PROPERTY cfgAlarmH : LREAL
GET
cfgAlarmH := _alarmH;
END_GET
SET
_alarmH := cfgAlarmH;
END_SET
END_PROPERTY

PROPERTY cfgAlarmHH : LREAL
GET
cfgAlarmHH := _alarmHH;
END_GET
SET
_alarmHH := cfgAlarmHH;
END_SET
END_PROPERTY

PROPERTY cfgAlarmL : LREAL
GET
cfgAlarmL := _alarmL;
END_GET
SET
_alarmL := cfgAlarmL;
END_SET
END_PROPERTY

PROPERTY cfgAlarmLL : LREAL
GET
cfgAlarmLL := _alarmLL;
END_GET
SET
_alarmLL := cfgAlarmLL;
END_SET
END_PROPERTY

PROPERTY cfgCalGain : LREAL
GET
cfgCalGain := _calGain;
END_GET
SET
_calGain := cfgCalGain;
END_SET
END_PROPERTY

PROPERTY cfgCalOffset : LREAL
GET
cfgCalOffset := _calOffset;
END_GET
SET
_calOffset := cfgCalOffset;
END_SET
END_PROPERTY

PROPERTY cfgEngUnit : STRING
GET
cfgEngUnit := _engUnit;
END_GET
SET
_engUnit := cfgEngUnit;
END_SET
END_PROPERTY

METHOD cmdReset : BOOL
setFault(0, '');
END_METHOD

METHOD PROTECTED FaultHandler : BOOL
VAR_INPUT
END_VAR
IF _alarmEnable THEN
	//L Warning
	_alarmDebounce[1](IN:=_alarmCooldown[1], PT:=T#30S);
	_alarmDebounce[2](IN:=_alarmCooldown[2], PT:=T#30S);
	IF _engValue < cfgAlarmL THEN
		IF NOT _alarmCooldown[1] THEN
			sendWarning(CONCAT(CONCAT('Low Warning - ', ANY_TO_STRING(TO_REAL(_engValue))),_EngUnit),1);
			_alarmCooldown[1] := TRUE;
		END_IF
	END_IF
	IF _alarmCooldown[1] AND _alarmDebounce[1].Q THEN
		_alarmCooldown[1] := FALSE;
	END_IF
	
	//H Warning
	IF _engValue > cfgAlarmH THEN
		IF NOT _alarmCooldown[2] THEN
			sendWarning(CONCAT(CONCAT('High Warning - ', ANY_TO_STRING(TO_REAL(_engValue))),_EngUnit),2);
			_alarmCooldown[2] := TRUE;
		END_IF
	END_IF
	IF _alarmCooldown[2] AND _alarmDebounce[2].Q THEN
		_alarmCooldown[2] := FALSE;
	END_IF
	
	IF _engValue < cfgAlarmLL THEN
		setFault(1,CONCAT(CONCAT('Low Alarm - ', ANY_TO_STRING(TO_REAL(_engValue))),_EngUnit));
	END_IF
	
	IF _engValue > cfgAlarmHH THEN
		setFault(1,CONCAT(CONCAT('High Alarm - ', ANY_TO_STRING(TO_REAL(_engValue))),_EngUnit));
	END_IF
	
	IF inpChannelDiag.error THEN
		setFault(1, 'Channel Error');
	END_IF
	
	IF inpChannelDiag.overrange THEN
		setFault(1, 'Overrange');
	END_IF
	
	IF inpChannelDiag.underrange THEN
		setFault(1, 'Underrange');
	END_IF
END_IF
END_METHOD

(*FB_Init is always available implicitly and it is used primarily for initialization.
The return value is not evaluated. For a specific influence, you can also declare the
methods explicitly and provide additional code there with the standard initialization
code. You can evaluate the return value.*)
METHOD FB_Init : BOOL
VAR_INPUT
	(* TRUE: the retain variables are initialized (reset warm / reset cold)*)
	bInitRetains	: BOOL;
	(* TRUE: the instance will be copied to the copy code afterward (online change)   *)
	bInCopyCode			: BOOL;
	cfgDeviceName		: STRING;
	cfgEnable			: BOOL;
	cfgInitEventClass	: BOOL;
	cfgAlarmEnable		: BOOL;
	cfgAlarmH			: LREAL;
	cfgAlarmHH			: LREAL;
	cfgAlarmL			: LREAL;
	cfgAlarmLL			: LREAL;
	cfgEngUnit			: STRING;
	cfgCalOffset		: LREAL;
	cfgCalGain			: LREAL := 1.0;	// omitted in the declaration = 1 (no correction)
END_VAR
THIS^.cfgDeviceName 		:= 		cfgDeviceName; 		
THIS^.cfgEnable 			:= 	    cfgEnable; 	
THIS^.cfgInitEventClass		:= 		cfgInitEventClass;
THIS^.cfgAlarmEnable		:=		cfgAlarmEnable;
THIS^.cfgAlarmH				:=		cfgAlarmH;
THIS^.cfgAlarmHH			:=		cfgAlarmHH;
THIS^.cfgAlarmL				:=		cfgAlarmL;
THIS^.cfgAlarmLL			:=		cfgAlarmLL;
THIS^.cfgCalOffset			:=		cfgCalOffset;
THIS^.cfgCalGain			:=		cfgCalGain;
THIS^.cfgEngUnit			:=		cfgEngUnit;

THIS^.HMI.cfgAlarmEnable	:= cfgAlarmEnable;
THIS^.HMI.cfgAlarmH			:= cfgAlarmH;
THIS^.HMI.cfgAlarmHH		:= cfgAlarmHH;
THIS^.HMI.cfgAlarmL			:= cfgAlarmL;
THIS^.HMI.cfgAlarmLL		:= cfgAlarmLL;
THIS^.HMI.cfgEngUnit		:= cfgEngUnit;
THIS^.HMI.cfgCalOffset		:= cfgCalOffset;
THIS^.HMI.cfgCalGain		:= cfgCalGain;
END_METHOD

METHOD scaleInput : BOOL
VAR_INPUT
END_VAR
IF cfgScalingNeeded THEN
	_sensorRawSignal	:= F_AnalogToEngUnit(inpRawIOChannel, cfgChannelMinInt, cfgChannelMaxInt, cfgSensorMin, cfgSensorMax);
	_engValue			:= (F_AnalogToEngUnit(stsSensorRawSignal, cfgSensorMin, cfgSensorMax, cfgEngUnitMin, cfgEngUnitMax) * _CalGain) + _CalOffset;
ELSE
	_sensorRawSignal := inpScaledIOChannel;
	_engValue		 := (inpScaledIOChannel * _CalGain) + _CalOffset;
END_IF
END_METHOD

METHOD PROTECTED setHMI : BOOL
VAR_INPUT
END_VAR
HMI.HMIbaseDevice := HMIbaseDevice;

HMI.stsEngValue 		:= _engValue;
HMI.stsSensorRawSignal	:= _sensorRawSignal;

cfgAlarmEnable		:= HMI.cfgAlarmEnable;
cfgAlarmH			:= HMI.cfgAlarmH;
cfgAlarmHH			:= HMI.cfgAlarmHH;
cfgAlarmL			:= HMI.cfgAlarmL;
cfgAlarmLL			:= HMI.cfgAlarmLL;
cfgCalOffset		:= HMI.cfgCalOffset;
cfgCalGain			:= HMI.cfgCalGain;
cfgEngUnit			:= HMI.cfgEngUnit;
END_METHOD

END_FUNCTION_BLOCK

// ---- POUs/FC/F_AnalogToEngUnit.TcPOU
FUNCTION F_AnalogToEngUnit : LREAL
VAR_INPUT
	inpRawSignal	:	LREAL;
	IO_min			:	LREAL;
	IO_max			: 	LREAL;
	engMin			:   LREAL;
	engMax			:	LREAL;
END_VAR

F_AnalogToEngUnit	:= engMin + (inpRawSignal - IO_min) * ((engmax - engmin) / (IO_max - IO_min));

END_FUNCTION

// ---- POUs/FBs/Devices/fb_Dev_AnalogSensor_Accelerometer.TcPOU
FUNCTION_BLOCK fb_Dev_AnalogSensor_Accelerometer EXTENDS fb_Dev_AnalogSensor

VAR_INPUT
	inpRawIOArray : ARRAY [0..49] OF INT;
END_VAR

VAR
	_mV_g : REAL;
	_engValueArray 			:  ARRAY [0..49] OF LREAL;
	_sensorRawSignalArray	:  ARRAY [0..49] OF LREAL;
END_VAR

VAR_OUTPUT
	stsSensorRawSignalArray	: ARRAY [0..49] OF LREAL;
	stsEngValueArray		: ARRAY [0..49] OF LREAL;
END_VAR

DeviceLogic();

scaleInput();

FaultHandler();

setHMI();

stsSensorRawSignalArray	:= _sensorRawSignalArray;
stsEngValueArray			:= _engValueArray;

(*FB_Init is always available implicitly and it is used primarily for initialization.
The return value is not evaluated. For a specific influence, you can also declare the
methods explicitly and provide additional code there with the standard initialization
code. You can evaluate the return value.*)
METHOD FB_Init : BOOL
VAR_INPUT
	(* TRUE: the retain variables are initialized (reset warm / reset cold)*)
	bInitRetains	: BOOL;
	(* TRUE: the instance will be copied to the copy code afterward (online change)   *)
bInCopyCode			: BOOL;
	cfgDeviceName		: STRING;
	cfgEnable			: BOOL;
	cfgInitEventClass	: BOOL;
	cfgAlarmEnable		: BOOL;
	cfgAlarmH			: LREAL;
	cfgAlarmHH			: LREAL;
	cfgAlarmL			: LREAL;
	cfgAlarmLL			: LREAL;
	cfgEngUnit			: STRING;
	cfgCalOffset		: LREAL;
	cfgCalGain			: LREAL := 1.0;	// omitted in the declaration = 1 (no correction)
	cfgmV_g				: REAL;
END_VAR
THIS^.cfgDeviceName 		:= 		cfgDeviceName; 		
THIS^.cfgEnable 			:= 	    cfgEnable; 	
THIS^.cfgInitEventClass		:= 		cfgInitEventClass;
THIS^.cfgAlarmEnable		:=		cfgAlarmEnable;
THIS^.cfgAlarmH				:=		cfgAlarmH;
THIS^.cfgAlarmHH			:=		cfgAlarmHH;
THIS^.cfgAlarmL				:=		cfgAlarmL;
THIS^.cfgAlarmLL			:=		cfgAlarmLL;
THIS^.cfgCalOffset			:=		cfgCalOffset;
THIS^.cfgCalGain			:=		cfgCalGain;
THIS^.cfgEngUnit			:=		cfgEngUnit;
THIS^._mV_g					:= 		cfgmV_g;

THIS^.HMI.cfgAlarmEnable	:= cfgAlarmEnable;
THIS^.HMI.cfgAlarmH			:= cfgAlarmH;
THIS^.HMI.cfgAlarmHH		:= cfgAlarmHH;
THIS^.HMI.cfgAlarmL			:= cfgAlarmL;
THIS^.HMI.cfgAlarmLL		:= cfgAlarmLL;
THIS^.HMI.cfgEngUnit		:= cfgEngUnit;
THIS^.HMI.cfgCalOffset		:= cfgCalOffset;
THIS^.HMI.cfgCalGain		:= cfgCalGain;
END_METHOD

PROPERTY mV_g : REAL
GET
mV_g := _mV_g;
END_GET
SET
_mV_g := mV_g;
END_SET
END_PROPERTY

METHOD scaleInput : BOOL
 VAR
	 i : INT;
 END_VAR
IF cfgScalingNeeded THEN
	FOR i := 0 TO 49 DO
		_sensorRawSignalArray[i]	:= F_AnalogToEngUnit(inpRawIOArray[i], cfgChannelMinInt, cfgChannelMaxInt, cfgSensorMin, cfgSensorMax);
		_engValueArray[i]			:= ((_sensorRawSignalArray[i]/_mV_g) * _CalGain) + _CalOffset;
	END_FOR
	
	
ELSE
	FOR i := 0 TO 49 DO
		_sensorRawSignalArray[i] := inpRawIOArray[i];
		_engValueArray[i]		 := (_sensorRawSignalArray[i] * _CalGain) + _CalOffset;
	END_FOR
END_IF
END_METHOD

END_FUNCTION_BLOCK

// ---- POUs/FBs/Devices/fb_Dev_AnalogSensor_CurrentTransducer.TcPOU
FUNCTION_BLOCK fb_Dev_AnalogSensor_CurrentTransducer EXTENDS fb_Dev_AnalogSensor
VAR_INPUT
END_VAR
VAR_OUTPUT
END_VAR
VAR
	_cfgShuntResValue	:LREAL;
	_cfgWindingRatio	:LREAL;
END_VAR

DeviceLogic();

scaleInput();

FaultHandler();

setHMI();

stsSensorRawSignal	:= _sensorRawSignal;
stsEngValue			:= _engValue;

PROPERTY cfgShuntResValue : LREAL
GET
cfgShuntResValue := _cfgShuntResValue;
END_GET
SET
_cfgShuntResValue := cfgShuntResValue;
END_SET
END_PROPERTY

PROPERTY cfgWindingRatio : LREAL
GET
cfgWindingRatio := _cfgWindingRatio;
END_GET
SET
_cfgWindingRatio := cfgWindingRatio;
END_SET
END_PROPERTY

(*FB_Init is always available implicitly and it is used primarily for initialization.
The return value is not evaluated. For a specific influence, you can also declare the
methods explicitly and provide additional code there with the standard initialization
code. You can evaluate the return value.*)
METHOD FB_Init : BOOL
VAR_INPUT
	(* TRUE: the retain variables are initialized (reset warm / reset cold)*)
	bInitRetains	: BOOL;
	(* TRUE: the instance will be copied to the copy code afterward (online change)   *)
	bInCopyCode	: BOOL;
	cfgDeviceName		: STRING;
	cfgEnable			: BOOL;
	cfgInitEventClass	: BOOL;
	cfgAlarmEnable		: BOOL;
	cfgAlarmH			: LREAL;
	cfgAlarmHH			: LREAL;
	cfgAlarmL			: LREAL;
	cfgAlarmLL			: LREAL;
	cfgEngUnit			: STRING;
	cfgCalOffset		: LREAL;
	cfgCalGain			: LREAL := 1.0;	// omitted in the declaration = 1 (no correction)
	cfgShuntResValue	: LREAL;
	cfgWindingRatio		: LREAL;
END_VAR
THIS^.cfgDeviceName 		:= 		cfgDeviceName; 		
THIS^.cfgEnable 			:= 	    cfgEnable; 	
THIS^.cfgInitEventClass		:= 		cfgInitEventClass;
THIS^.cfgAlarmEnable		:=		cfgAlarmEnable;
THIS^.cfgAlarmH				:=		cfgAlarmH;
THIS^.cfgAlarmHH			:=		cfgAlarmHH;
THIS^.cfgAlarmL				:=		cfgAlarmL;
THIS^.cfgAlarmLL			:=		cfgAlarmLL;
THIS^.cfgCalOffset			:=		cfgCalOffset;
THIS^.cfgCalGain			:=		cfgCalGain;
THIS^.cfgEngUnit			:=		cfgEngUnit;
THIS^.cfgShuntResValue		:=		cfgShuntResValue;
THIS^.cfgWindingRatio		:=		cfgWindingRatio;

THIS^.HMI.cfgAlarmEnable	:= cfgAlarmEnable;
THIS^.HMI.cfgAlarmH			:= cfgAlarmH;
THIS^.HMI.cfgAlarmHH		:= cfgAlarmHH;
THIS^.HMI.cfgAlarmL			:= cfgAlarmL;
THIS^.HMI.cfgAlarmLL		:= cfgAlarmLL;
THIS^.HMI.cfgEngUnit		:= cfgEngUnit;
THIS^.HMI.cfgCalOffset		:= cfgCalOffset;
THIS^.HMI.cfgCalGain		:= cfgCalGain;
END_METHOD

METHOD scaleInput : BOOL
IF cfgScalingNeeded THEN
	_sensorRawSignal	:= F_AnalogToEngUnit(inpRawIOChannel, cfgChannelMinInt, cfgChannelMaxInt, cfgSensorMin, cfgSensorMax);
	_engValue			:= (_sensorRawSignal * _cfgWindingRatio / _cfgShuntResValue) * _CalGain + _calOffset;
ELSE
	_sensorRawSignal := inpRawIOChannel;
	_engValue		 := (inpRawIOChannel * _CalGain) + _calOffset;
END_IF
END_METHOD

END_FUNCTION_BLOCK

// ---- POUs/FBs/Devices/fb_Dev_AnalogSensor_ELM_10x.TcPOU
FUNCTION_BLOCK fb_Dev_AnalogSensor_ELM_10x EXTENDS fb_Dev_AnalogSensor
VAR_INPUT
	inpRawIOChannelArray			: ARRAY [1..10] OF DINT;
END_VAR
VAR_OUTPUT
	stsSensorRawSignalArray	: ARRAY [1..10] OF LREAL;
	stsEngValueArray		: ARRAY [1..10] OF LREAL;
	stsEngValueRMS			: LREAL;
END_VAR
VAR
	_sensorRawSignalArray			: ARRAY [1..10] OF LREAL;
	_engValueArray					: ARRAY [1..10] OF LREAL;
	_engValueRMS					: LREAL;
END_VAR

// This FB is intended for a ELM IO card set to 10x overscan with a 1ms CPU cycletime

DeviceLogic();

scaleInput();

FaultHandler();

setHMI();

stsSensorRawSignalArray		:= _sensorRawSignalArray;
stsEngValueArray			:= _engValueArray;

stsSensorRawSignal 			:= _sensorRawSignal;
stsEngValue					:= _engValue;

METHOD scaleInput : BOOL
VAR
	i : INT;
	tempRaw : LREAL := 0.0;
	tempEng : LREAL := 0.0;
	tempEngSqSum 	: LREAL := 0.0;
END_VAR
FOR i := 1 TO 10 DO
	_sensorRawSignalArray[i]	:= F_AnalogToEngUnit(inpRawIOChannelArray[i], cfgChannelMinInt, cfgChannelMaxInt, cfgSensorMin, cfgSensorMax);
	_engValueArray[i]			:= (F_AnalogToEngUnit(_sensorRawSignalArray[i], cfgSensorMin, cfgSensorMax, cfgEngUnitMin, cfgEngUnitMax) * _CalGain) + _CalOffset;
	tempRaw := tempRaw + _sensorRawSignalArray[i];
	tempEng := tempEng + _engValueArray[i];
	tempEngSqSum := tempEngSqSum + _engValueArray[i] * _engValueArray[i];
END_FOR

_sensorRawSignal	:= tempRaw / 10;
_engValue			:= tempEng / 10;
_engValueRMS		:= SQRT(tempEngSqSum / 10);
END_METHOD

END_FUNCTION_BLOCK

// ---- POUs/FBs/Devices/fb_Dev_AnalogSensor_ELM_10x_CurrentTransducer.TcPOU
FUNCTION_BLOCK fb_Dev_AnalogSensor_ELM_10x_CurrentTransducer EXTENDS fb_Dev_AnalogSensor_CurrentTransducer
VAR_INPUT
	inpRawIOChannelArray			: ARRAY [1..10] OF DINT;
END_VAR
VAR_OUTPUT
	stsSensorRawSignalArray	: ARRAY [1..10] OF LREAL;
	stsEngValueArray		: ARRAY [1..10] OF LREAL;
	stsEngValueRMS			: LREAL;
END_VAR
VAR
	_sensorRawSignalArray			: ARRAY [1..10] OF LREAL;
	_engValueArray					: ARRAY [1..10] OF LREAL;
	_engValueRMS					: LREAL;
END_VAR

// This FB is intended for a ELM IO card set to 10x overscan with a 1ms CPU cycletime

DeviceLogic();

scaleInput();

FaultHandler();

setHMI();

stsSensorRawSignalArray		:= _sensorRawSignalArray;
stsEngValueArray			:= _engValueArray;

stsSensorRawSignal 			:= _sensorRawSignal;
stsEngValue					:= _engValue;
stsEngValueRMS				:= _engValueRMS;

METHOD scaleInput : BOOL
VAR
	i : INT;
	tempRaw 		: LREAL := 0.0;
	tempEng 		: LREAL := 0.0;
	tempEngSqSum 	: LREAL := 0.0;
END_VAR
FOR i := 1 TO 10 DO
	_sensorRawSignalArray[i]	:= F_AnalogToEngUnit(inpRawIOChannelArray[i], cfgChannelMinInt, cfgChannelMaxInt, cfgSensorMin, cfgSensorMax);
	_engValueArray[i]			:= (_sensorRawSignalArray[i] * _cfgWindingRatio / _cfgShuntResValue) * _CalGain + _calOffset;
	tempRaw := tempRaw + _sensorRawSignalArray[i];
	tempEng := tempEng + _engValueArray[i];
	tempEngSqSum := tempEngSqSum + _engValueArray[i] * _engValueArray[i];
	
END_FOR

_sensorRawSignal	:= tempRaw / 10;
_engValue			:= tempEng / 10;
_engValueRMS		:= SQRT(tempEngSqSum / 10);
END_METHOD

END_FUNCTION_BLOCK

// ---- POUs/FBs/Devices/fb_Dev_ControlValve_Modulating_INT.TcPOU
FUNCTION_BLOCK fb_Dev_ControlValve_Modulating_INT
VAR_INPUT
	IO_valveFeedback	: INT;
	IO_valveOutput		: POINTER TO INT;
	inpAuto				: BOOL;
	inpReset			: BOOL;
	inpInterlockBypass	: BOOL;
	faultMonitor		: POINTER TO fb_FaultMonitor;
END_VAR

VAR
	valveFeedback_scaled	: LREAL;
	valveFeedback_volts		: LREAL;
	_valveName				: STRING;
	Valve					: fb_Dev_ControlValve_Modulating(cfgDeviceName := _valveName, cfgEnable := TRUE, cfgInitEventClass := TRUE);
	_valvePositionCmd		: LREAL;
	_valveOutput_volts		: LREAL;
	
END_VAR
VAR_OUTPUT
	outValvePosition	: LREAL;
	stsValveFeedback	: LREAL;
END_VAR

//INPUTS AND OUTPUTS FOR THIS FB VARIANT ARE UNSCALLED ANALOG VALUES
valveFeedback_volts	:=  F_AnalogToEngUnit(TO_REAL(IO_valveFeedback), -32767, 32767, -10, 10);
valveFeedback_scaled := F_AnalogToEngUnit(valveFeedback_volts, 2, 10, 0, 100);

Valve(inpAuto := inpAuto, inpReset := inpReset, inpInterlockBypass := inpInterlockBypass, faultMonitor:=faultMonitor
		, inpValvePosition := valveFeedback_scaled);
		
outValvePosition := Valve.outValvePosition;
stsValveFeedback := Valve.stsValveFeedback;

Valve.valvePosition := _valvePositionCmd;

_valveOutput_volts := F_AnalogToEngUnit(Valve.outValvePosition, 0, 100, 2, 10);	
IO_valveOutput^ := TO_INT(F_AnalogToEngUnit(inpRawSignal := _valveOutput_volts, IO_min := -10, IO_max := 10, engMin := -32767, engMax := 32767));

PROPERTY cmdSetValvePosition : LREAL
SET
_valvePositionCmd := cmdSetValvePosition;
END_SET
END_PROPERTY

//FB_Init is always available implicitly and it is used primarily for initialization.
//The return value is not evaluated. For a specific influence, you can also declare the
//methods explicitly and provide additional code there with the standard initialization
//code. You can evaluate the return value.
METHOD FB_Init: BOOL
VAR_INPUT
    bInitRetains	: BOOL; // TRUE: the retain variables are initialized (reset warm / reset cold)
    bInCopyCode		: BOOL;  // TRUE: the instance will be copied to the copy code afterward (online change) 
	cfgDeviceName	: STRING;  
	cfgInitPosition  : LREAL;
END_VAR
THIS^._valveName 			:= cfgDeviceName;
THIS^.Valve.cfgDeviceName 	:= cfgDeviceName;
THIS^.cmdSetValvePosition   := cfgInitPosition;
END_METHOD

END_FUNCTION_BLOCK

// ---- POUs/FBs/Devices/fb_Dev_ControlValve_Modulating.TcPOU
FUNCTION_BLOCK fb_Dev_ControlValve_Modulating EXTENDS abs_fb_Device
VAR_INPUT
	inpValvePosition	: LREAL;
END_VAR

VAR
	transMantoAuto	: R_TRIG;
	transAutoToMan	: F_TRIG;
END_VAR

VAR PERSISTENT
	HMI				: ST_ControlValve_Modulating_HMI_Interface;
	_valvePosition	: LREAL;
END_VAR


VAR_OUTPUT
	outValvePosition	: LREAL;
	stsValveFeedback	: LREAL;
END_VAR

DeviceLogic();
Interlock.name := _DeviceName;
Interlock(inpConfig := _dataInterlock);

faultHandler();

transManToAuto(CLK:=_inAuto);
transAutoToMan(CLK:=_inAuto);

stsValveFeedback := inpValvePosition;

// Maintain valve position during man/auto machine state changes
IF transManToAuto.Q THEN
	_valvePosition := HMI.ocmdValvePosition;
END_IF

IF transAutoToMan.Q THEN
	HMI.ocmdValvePosition := _valvePosition;
END_IF

IF NOT stsFaulted AND Interlock.outInterlockOK THEN
	IF _inAuto THEN
		outValvePosition := _valvePosition;
	ELSE
		outValvePosition := HMI.ocmdValvePosition;
	END_IF
END_IF

HMI.stsValveFeedback := stsValveFeedback;
HMI.stsValvePosition := outValvePosition;
HMI.HMIbaseDevice := HMIBaseDevice;

METHOD faultHandler : BOOL
VAR_INPUT
END_VAR
IF stsValveFeedback < -1 AND _warnChannels[1] = '' THEN
	sendWarning('Valve feedback not present', 1);
END_IF
END_METHOD

PROPERTY valvePosition : LREAL
GET
valvePosition := _valvePosition;
END_GET
SET
_valvePosition := valvePosition;
END_SET
END_PROPERTY

END_FUNCTION_BLOCK

// ---- POUs/FBs/Devices/fb_Dev_Pump_ABBACS580.TcPOU
FUNCTION_BLOCK fb_Dev_Pump_ABBACS580 EXTENDS abs_fb_Device
VAR_INPUT
	inpESTOPs_OK			: BOOL;		// 1 = ESTOPs healthy, 0 = ESTOP active
	inpMachineSTOP			: BOOL;
	inpOverpressureTrip		: BOOL;		// asserted by caller when pressure > limit
END_VAR

VAR PERSISTENT
	HMI						: ST_Pump_ABBACS580_HMI_Interface;
END_VAR

VAR
	// Embedded VFD driver (forward-only operation enforced by this wrapper)
	VFD : fb_Dev_VFD_ABBACS580(
		cfgDeviceName		:= CONCAT(_deviceName, ' VFD'),
		cfgEnable			:= TRUE,
		cfgInitEventClass	:= TRUE,
		cfgIPAddress		:= _ipAddress,
		cfgUnitID			:= _unitId);

	// Pump-level control state (set by cmdRun / cmdSetpoint in auto mode,
	// sourced from VFD.HMI in manual mode)
	_ctrlRun				: BOOL;
	_ctrlSetpoint			: LREAL;	// 0..100 percent
	_resetTrig				: R_TRIG;

	// Modbus addressing mirrors (set via cfg* properties before enable)
	_ipAddress				: STRING(15) := '192.168.1.50';
	_unitId					: BYTE := 1;

	// Trip bit OR'd into the VFD's outbound CW
	_trippedBitMask			: WORD;

	// Interlock array
	_interlocks				: ARRAY[1..10] OF BOOL;
END_VAR

VAR_OUTPUT
	stsOverpressureTripped	: BOOL;
END_VAR

DeviceLogic();

// Propagate Modbus addressing into the inner VFD. Required because TwinCAT
// initializes embedded FBs in VAR declaration order: VFD.FB_Init runs before
// _ipAddress is default-initialized AND before pump.FB_Init applies any
// override, so VFD._ipAddress would otherwise be locked at empty. Assigning
// each scan is cheap and is consumed once by VFD's one-shot _modbusInit.
VFD.cfgIPAddress	:= _ipAddress;
VFD.cfgUnitID		:= _unitId;

// Continuous trip bit. Drive will fault via External event 1 IF par 31.01
// has been configured on the drive (e.g. to FBA Main CW bit 12).
IF inpOverpressureTrip THEN
	_trippedBitMask := 16#1000;
ELSE
	_trippedBitMask := 16#0000;
END_IF
stsOverpressureTripped := inpOverpressureTrip;

// Manual mode: source commands from pump HMI. Forward-only is enforced by the
// pump's BOOL ocmdRun and 0..100 setpoint clamp — the inner VFD never sees a
// reverse command because we force it to auto mode below.
IF _enabled THEN
	IF NOT _inAuto THEN
		_ctrlRun		:= HMI.ocmdRun;
		_ctrlSetpoint	:= LIMIT(0.0, HMI.ocmdSetpoint, 100.0);
	END_IF
END_IF

_resetTrig(CLK := HMI.ocmdReset);
IF _resetTrig.Q THEN
	cmdReset();
END_IF

// Pump-level interlocks
_interlocks[1] := inpESTOPs_OK;
cmdSetInterlock(1, 'ESTOPs OK', _interlocks[1]);

_interlocks[2] := NOT inpMachineSTOP;
cmdSetInterlock(2, 'Machine STOP Not Active', _interlocks[2]);

_interlocks[3] := NOT inpOverpressureTrip;
cmdSetInterlock(3, 'Pressure below limit', _interlocks[3]);

FaultHandler();

// Interlock enforcement (force stop on broken interlock; mirror to pump HMI
// so the operator sees the run command drop)
IF NOT interlock.outInterlockOK THEN
	_ctrlRun	:= FALSE;
	HMI.ocmdRun	:= FALSE;
END_IF

// Drive the inner VFD with the forward-only API.
// inpAuto is forced TRUE so VFD never sources commands from its own HMI —
// pump HMI is the sole operator surface. cmdEnable / cmdSetpoint are the
// single source of truth for the inner VFD.
IF _ctrlRun THEN
	VFD.cmdEnable(1);
ELSE
	VFD.cmdEnable(0);
END_IF
VFD.cmdSetpoint(_ctrlSetpoint);

VFD(
	inpAuto				:= TRUE,
	inpReset			:= inpReset,
	inpInterlockBypass	:= inpInterlockBypass,
	inpESTOPs_OK		:= inpESTOPs_OK,
	inpMachineSTOP		:= inpMachineSTOP,
	inpCWAuxBitMask		:= _trippedBitMask);

updateHMI();

PROPERTY cfgIPAddress : STRING(15)
GET
cfgIPAddress := _ipAddress;
END_GET
SET
_ipAddress := cfgIPAddress;
END_SET
END_PROPERTY

PROPERTY cfgUnitID : BYTE
GET
cfgUnitID := _unitId;
END_GET
SET
_unitId := cfgUnitID;
END_SET
END_PROPERTY

METHOD PUBLIC cmdRun : BOOL
VAR_INPUT
	command		: BOOL;		// TRUE = run forward, FALSE = stop
END_VAR
_ctrlRun := command;
END_METHOD

METHOD PUBLIC cmdSetpoint : BOOL
VAR_INPUT
	setpoint	: LREAL;	// 0..100 percent (negative clamped to 0)
END_VAR
_ctrlSetpoint := LIMIT(0.0, setpoint, 100.0);
END_METHOD

METHOD PUBLIC cmdReset : BOOL
setFault(0, '');
VFD.cmdReset();
END_METHOD

METHOD PRIVATE FaultHandler : BOOL
VAR_INPUT
END_VAR
// Overpressure: latch as a pump fault so the operator sees what stopped the
// pump. Without this, the interlock-3 enforcement above silently force-stops
// the pump with no fault state.
IF inpOverpressureTrip THEN
	setFault(1, 'Overpressure trip');
END_IF

// Forward drive-level trip as a pump fault. Evaluated after overpressure so
// that if both fire simultaneously, the drive fault code surfaces in the
// description (overpressure already routed to the drive via CW bit 12).
IF VFD.stsTripped THEN
	setFault(1, CONCAT('VFD Tripped, code ', UINT_TO_STRING(VFD.stsFaultCode)));
END_IF

// Drive-level warning passthrough
IF VFD.stsAlarm THEN
	sendWarning('Drive alarm active', 10);
END_IF
END_METHOD

METHOD PRIVATE updateHMI : BOOL
VAR
END_VAR
HMI.HMIbaseDevice			:= HMIbaseDevice;
HMI.stsInterlocks			:= interlock.getHMIdata();
HMI.stsOverpressureTripped	:= stsOverpressureTripped;
END_METHOD

METHOD FB_Init : BOOL
VAR_INPUT
	bInitRetains		: BOOL;
	bInCopyCode			: BOOL;
	cfgDeviceName		: STRING;
	cfgEnable			: BOOL;
	cfgInitEventClass	: BOOL;
	cfgIPAddress		: STRING(15);
	cfgUnitID			: BYTE;
END_VAR
THIS^.cfgDeviceName		:= cfgDeviceName;
THIS^.cfgEnable			:= cfgEnable;
THIS^.cfgInitEventClass	:= cfgInitEventClass;
THIS^.cfgIPAddress		:= cfgIPAddress;
THIS^.cfgUnitID			:= cfgUnitID;
END_METHOD

END_FUNCTION_BLOCK

// ---- POUs/FBs/Devices/fb_Dev_VFD_ABBACS580.TcPOU
FUNCTION_BLOCK fb_Dev_VFD_ABBACS580 EXTENDS abs_fb_Device
VAR_INPUT
	inpESTOPs_OK		: BOOL;		// 1 = ESTOPs healthy, 0 = ESTOP active
	inpMachineSTOP		: BOOL;
	inpCWAuxBitMask		: WORD;		// OR'd into outbound CW (app-specific bits 12-15)
END_VAR

VAR PERSISTENT
	HMI					: ST_VFD_ABBACS580_HMI_Interface;
END_VAR

VAR
	// Embedded Modbus TCP client
	_modbus				: fb_Modbus_Driver;
	_modbusInit			: BOOL;

	// Read signal config.
	// SW + ACT1 come from the cyclic data exchange (regs 40004/40005, fixed by
	// ABB Drives Classic profile). Everything else uses direct parameter access
	// (register = 40000 + group*100 + index) so no drive-side slot mapping
	// configuration (par 52.04+, refresh) is required. The driver issues
	// multiple non-contiguous FC03 transactions per poll cycle; latency is
	// dominated by the cyclic SW/ACT1 reads regardless.
	_arrReadConfig		: ARRAY[1..8] OF ST_MBSignalConfig := [
		(modbusAddr := 40004, dataType := E_MBDataType.mbUInt16, tag := 'SW'),			// cyclic
		(modbusAddr := 40005, dataType := E_MBDataType.mbInt16,  tag := 'ACT1'),		// cyclic
		(modbusAddr := 40107, dataType := E_MBDataType.mbUInt16, tag := 'MotorCurrent'),// par 01.07 direct
		(modbusAddr := 40111, dataType := E_MBDataType.mbUInt16, tag := 'DCBus'),		// par 01.11 direct
		(modbusAddr := 40106, dataType := E_MBDataType.mbInt16,  tag := 'OutFreq'),		// par 01.06 direct
		(modbusAddr := 40110, dataType := E_MBDataType.mbInt16,  tag := 'Torque'),		// par 01.10 direct
		(modbusAddr := 40511, dataType := E_MBDataType.mbUInt16, tag := 'InvTemp'),		// par 05.11 direct
		(modbusAddr := 40411, dataType := E_MBDataType.mbUInt16, tag := 'FaultCode')];	// par 04.11 direct
	_arrReadResults		: ARRAY[1..8] OF ST_MBReadResult;

	// Write signal config: CW + REF1 (contiguous => single FC16)
	_arrWriteConfig		: ARRAY[1..2] OF ST_MBSignalConfig := [
		(modbusAddr := 40001, dataType := E_MBDataType.mbUInt16, tag := 'CW'),
		(modbusAddr := 40002, dataType := E_MBDataType.mbInt16,  tag := 'REF1')];
	_arrWriteData		: ARRAY[1..2] OF ST_MBWriteData;

	// Application-level control signals
	_ctrlRunMode		: USINT;		// 0=stop, 1=fwd, 2=reverse
	_ctrlSetpoint		: LREAL;		// -100..+100 percent
	_resetTrig			: R_TRIG;

	// Event-logging edge detection
	_lastLoggedRunMode	: USINT;
	_lastLoggedSetpoint	: LREAL;
	_trippedTrig		: R_TRIG;

	// CW state machine
	_cwState			: INT;			// 0=Idle, 1=Running, 2=FaultPending, 3=ResetSequence
	_cwCurrent			: WORD := 16#047E;	// init 1150 (Ready) so first write is benign
	_resetTimeout		: TON;
	_readyTimeout		: TON;
	_safetyStopActive	: BOOL;

	// Parsed status word
	_swRaw				: WORD;
	_stsRdyOn			: BOOL;
	_stsRdyRun			: BOOL;
	_stsRunning			: BOOL;
	_stsTripped			: BOOL;
	_stsAlarm			: BOOL;
	_stsAtSetpoint		: BOOL;
	_stsRemote			: BOOL;
	_stsSwOnInhibit		: BOOL;

	// Engineering-unit telemetry
	_telemetry			: ST_VFD_ABBACS580_Telemetry;
	_stateString		: STRING;

	// Interlock array (parallels Pump_SPAL pattern)
	_interlocks			: ARRAY[1..10] OF BOOL;

	// Modbus configuration mirrors (set via cfg* properties before enable)
	_ipAddress			: STRING(15) := '192.168.1.50';
	_unitId				: BYTE := 1;
END_VAR

VAR_OUTPUT
	stsRunning			: BOOL;
	stsReady			: BOOL;
	stsAtSetpoint		: BOOL;
	stsRemote			: BOOL;
	stsAlarm			: BOOL;
	stsTripped			: BOOL;
	stsActualSpeed		: LREAL;	// percent
	stsActualCurrent	: LREAL;	// A
	stsActualTorque	: LREAL;		// %
	stsOutputFreq		: LREAL;	// Hz, signed
	stsDCBusVoltage	: LREAL;		// VDC
	stsInverterTemp	: LREAL;		// %
	stsFaultCode		: UINT;	// 0 unless drive is actively tripped
	stsFaultText		: STRING;	// decoded fault name; empty unless tripped
	stsCommsConnected	: BOOL;
END_VAR

DeviceLogic();

// One-time Modbus driver configuration (properties lock after _initialized := TRUE)
IF NOT _modbusInit THEN
	_modbus.ipAddress				:= _ipAddress;
	_modbus.unitId					:= _unitId;
	_modbus.port					:= 502;
	_modbus.timeout					:= T#500MS;
	_modbus.pollInterval			:= T#50MS;
	_modbus.writeCycleInterval		:= T#100MS;
	_modbus.wordOrder				:= E_WordOrder.BigEndian;
	_modbus.maxConsecFails			:= 3;
	_modbus.reconnectDelay			:= T#2S;
	_modbus.maxReconnectAttempts	:= 10;
	_modbus.staleThreshold			:= T#2S;
	_modbus.readSignalCount			:= 8;
	_modbus.writeSignalCount		:= 2;
	_modbusInit := TRUE;
END_IF

// Drive the embedded Modbus client
_modbus(
	inpEnable			:= _enabled,
	inpPtrReadConfig	:= ADR(_arrReadConfig),
	inpPtrWriteConfig	:= ADR(_arrWriteConfig),
	inpPtrReadResults	:= ADR(_arrReadResults),
	inpPtrWriteData		:= ADR(_arrWriteData));
_modbus.cycle();

parseDriveFeedback();

// Interlocks (numbered like Pump_SPAL)
_interlocks[1] := inpESTOPs_OK;
cmdSetInterlock(1, 'ESTOPs OK', _interlocks[1]);

_interlocks[2] := NOT inpMachineSTOP;
cmdSetInterlock(2, 'Machine STOP Not Active', _interlocks[2]);

_interlocks[3] := _modbus.stsStatus.connected AND NOT _modbus.stsStatus.faulted;
cmdSetInterlock(3, 'Modbus comms OK', _interlocks[3]);

_interlocks[4] := _stsRemote;
cmdSetInterlock(4, 'Drive in Remote mode', _interlocks[4]);

_safetyStopActive := (NOT inpESTOPs_OK) OR inpMachineSTOP;

// HMI command surface — only honoured in manual mode (parallels Pump_SPAL)
IF _enabled THEN
	IF NOT _inAuto THEN
		_ctrlRunMode	:= HMI.ocmdRunMode;
		_ctrlSetpoint	:= HMI.ocmdSetpoint;
	END_IF
END_IF

_resetTrig(CLK := HMI.ocmdReset);
IF _resetTrig.Q THEN
	cmdReset();
END_IF

FaultHandler();

// Interlock enforcement: force commanded mode to stop if broken.
// (Coast-vs-ramp routing happens inside controlWordSequencer via _safetyStopActive.)
IF NOT interlock.outInterlockOK THEN
	_ctrlRunMode	:= 0;
	HMI.ocmdRunMode	:= 0;
END_IF

controlWordSequencer();

// Marshal CW + REF1 into Modbus write buffers
// inpCWAuxBitMask lets a wrapper FB inject app-specific bits (e.g. CW bit 12 for external-event trip)
_arrWriteData[1].valueUint	:= WORD_TO_UINT(_cwCurrent OR inpCWAuxBitMask);
_arrWriteData[2].valueInt	:= LREAL_TO_INT(LIMIT(-100.0, _ctrlSetpoint, 100.0) * 200.0);

// Event-based logging (run mode change, setpoint change, fault entry)
IF _ctrlRunMode <> _lastLoggedRunMode THEN
	CASE _ctrlRunMode OF
		0:	sendLog('Stop command', 1);
		1:	sendLog(CONCAT('Run forward @ ', LREAL_TO_STRING(_ctrlSetpoint)), 1);
		2:	sendLog(CONCAT('Run reverse @ ', LREAL_TO_STRING(_ctrlSetpoint)), 1);
	END_CASE
	_lastLoggedRunMode := _ctrlRunMode;
END_IF

IF ABS(_ctrlSetpoint - _lastLoggedSetpoint) >= 0.1 THEN
	sendLog(CONCAT('Setpoint = ', LREAL_TO_STRING(_ctrlSetpoint)), 2);
	_lastLoggedSetpoint := _ctrlSetpoint;
END_IF

_trippedTrig(CLK := _stsTripped);
IF _trippedTrig.Q THEN
	sendLog(CONCAT('Drive tripped, fault code ', UINT_TO_STRING(_telemetry.faultCode)), 3);
END_IF

updateHMI();

// Public outputs
stsRunning			:= _stsRunning;
stsReady			:= _stsRdyOn AND _stsRdyRun;
stsAtSetpoint		:= _stsAtSetpoint;
stsRemote			:= _stsRemote;
stsAlarm			:= _stsAlarm;
stsTripped			:= _stsTripped;
stsActualSpeed		:= _telemetry.actualSpeed;
stsActualCurrent	:= _telemetry.motorCurrent;
stsActualTorque		:= _telemetry.motorTorque;
stsOutputFreq		:= _telemetry.outputFreq;
stsDCBusVoltage		:= _telemetry.dcBusVoltage;
stsInverterTemp		:= _telemetry.inverterTemp;
// Gate fault code & decoded text by active trip. Par 04.11 latches the LAST
// fault on the drive even after a reset, which is misleading on the HMI when
// the drive isn't actually faulted.
IF _stsTripped THEN
	stsFaultCode	:= _telemetry.faultCode;
	stsFaultText	:= decodeFaultCode(_telemetry.faultCode);
ELSE
	stsFaultCode	:= 0;
	stsFaultText	:= '';
END_IF
// AND-ing with signal quality so this agrees with the 'No Comms' branch in
// parseDriveFeedback. The driver's 'connected' flag lags reality (tracks
// TCP / driver state, only drops after maxConsecFails retries), while signal
// quality flips on the first failed read. Operator-facing status should
// reflect data freshness, not socket state.
stsCommsConnected	:= _modbus.stsStatus.connected AND (_arrReadResults[1].quality = E_SignalQuality.Good);

PROPERTY cfgIPAddress : STRING(15)
GET
cfgIPAddress := _ipAddress;
END_GET
SET
_ipAddress := cfgIPAddress;
END_SET
END_PROPERTY

PROPERTY cfgUnitID : BYTE
GET
cfgUnitID := _unitId;
END_GET
SET
_unitId := cfgUnitID;
END_SET
END_PROPERTY

METHOD PUBLIC cmdEnable : BOOL
VAR_INPUT
	command		: USINT;	// 0=stop, 1=run forward, 2=run reverse
END_VAR
IF command <= 2 THEN
	_ctrlRunMode := command;
END_IF
END_METHOD

METHOD PUBLIC cmdSetpoint : BOOL
VAR_INPUT
	setpoint	: LREAL;	// percent, -100..+100
END_VAR
_ctrlSetpoint := LIMIT(-100.0, setpoint, 100.0);
END_METHOD

METHOD PUBLIC cmdReset : BOOL
setFault(0, '');
IF _stsTripped THEN
	_cwState := 3;
END_IF
// A driver that gave up after maxReconnectAttempts restarts on reset (it no longer needs a
// PLC restart to recover).
IF _modbus.stsStatus.faulted THEN
	_modbus.cmdReset();
END_IF
END_METHOD

METHOD PRIVATE controlWordSequencer : BOOL
VAR_INPUT
END_VAR
// CW values per abbmodbus.md section 3:
//   16#047E (1150) = Ready / ramp-stop
//   16#047D (1149) = Coast stop (OFF2)
//   16#047F (1151) = Run forward
//   16#0C7F (3199) = Run reverse
//   16#04FF (1279) = Fault reset (CW.bit7 high)

CASE _cwState OF
	0:	// Idle / Ready
		IF _safetyStopActive THEN
			_cwCurrent := 16#047D;		// coast on safety interlock
		ELSE
			_cwCurrent := 16#047E;		// normal ramp stop / ready
		END_IF
		_readyTimeout(IN := _ctrlRunMode > 0, PT := T#10S);
		// RDY_RUN (SW bit 1) is a consequence of releasing OFF1 (CW bit 0 -> 1),
		// not a precondition. Gating on it deadlocks the drive in
		// READY_TO_SWITCH_ON. RDY_ON alone is the correct precondition.
		IF _ctrlRunMode > 0
		   AND _stsRdyOn
		   AND NOT _stsTripped
		   AND NOT _safetyStopActive THEN
			_cwState := 1;
			_readyTimeout(IN := FALSE);
		ELSIF _readyTimeout.Q THEN
			setFault(1, 'Drive did not reach Ready within 10s');
			_readyTimeout(IN := FALSE);
		END_IF

	1:	// Running
		IF _stsTripped THEN
			_cwState := 2;
		ELSIF _ctrlRunMode = 0 OR _safetyStopActive THEN
			_cwState := 0;
		ELSIF _ctrlRunMode = 1 THEN
			_cwCurrent := 16#047F;		// run forward
		ELSIF _ctrlRunMode = 2 THEN
			_cwCurrent := 16#0C7F;		// run reverse
		END_IF

	2:	// FaultPending — wait for reset
		_cwCurrent := 16#047E;
		IF NOT _stsTripped THEN
			_cwState := 0;
		END_IF

	3:	// ResetSequence — hold 1279 until SW.bit3 deasserts (max 3s)
		_cwCurrent := 16#04FF;
		_resetTimeout(IN := TRUE, PT := T#3S);
		IF NOT _stsTripped THEN
			_cwState := 0;
			_resetTimeout(IN := FALSE);
		ELSIF _resetTimeout.Q THEN
			setFault(1, 'Fault reset did not clear after 3s');
			_cwState := 2;
			_resetTimeout(IN := FALSE);
		END_IF
END_CASE
END_METHOD

METHOD PRIVATE parseDriveFeedback : BOOL
VAR_INPUT
END_VAR
// SW (par 58.104 default mapping)
IF _arrReadResults[1].quality = E_SignalQuality.Good THEN
	_swRaw			:= UINT_TO_WORD(_arrReadResults[1].valueUint);
	_stsRdyOn		:= (_swRaw AND 16#0001) <> 0;	// bit 0 RDY_ON
	_stsRdyRun		:= (_swRaw AND 16#0002) <> 0;	// bit 1 RDY_RUN
	_stsRunning		:= (_swRaw AND 16#0004) <> 0;	// bit 2 RDY_REF (operation enabled)
	_stsTripped		:= (_swRaw AND 16#0008) <> 0;	// bit 3 TRIPPED
	_stsSwOnInhibit	:= (_swRaw AND 16#0040) <> 0;	// bit 6 SWC_ON_INHIB
	_stsAlarm		:= (_swRaw AND 16#0080) <> 0;	// bit 7 ALARM
	_stsAtSetpoint	:= (_swRaw AND 16#0100) <> 0;	// bit 8 AT_SETPOINT
	_stsRemote		:= (_swRaw AND 16#0200) <> 0;	// bit 9 REMOTE
END_IF

// ACT1: -20000..+20000 = -100..+100%
IF _arrReadResults[2].quality = E_SignalQuality.Good THEN
	_telemetry.actualSpeed	:= INT_TO_LREAL(_arrReadResults[2].valueInt) / 200.0;
END_IF

// Motor current (par 01.07, default whole A)
IF _arrReadResults[3].quality = E_SignalQuality.Good THEN
	_telemetry.motorCurrent	:= UINT_TO_LREAL(_arrReadResults[3].valueUint);
END_IF

// DC bus voltage (par 01.11, raw 0.1 VDC)
IF _arrReadResults[4].quality = E_SignalQuality.Good THEN
	_telemetry.dcBusVoltage	:= UINT_TO_LREAL(_arrReadResults[4].valueUint) / 10.0;
END_IF

// Output frequency (par 01.06, raw -20000..+20000 = -100..+100% of par 46.02)
IF _arrReadResults[5].quality = E_SignalQuality.Good THEN
	_telemetry.outputFreq	:= INT_TO_LREAL(_arrReadResults[5].valueInt) * 60.0 / 20000.0;
END_IF

// Motor torque (par 01.10, raw 0.01%)
IF _arrReadResults[6].quality = E_SignalQuality.Good THEN
	_telemetry.motorTorque	:= INT_TO_LREAL(_arrReadResults[6].valueInt) / 100.0;
END_IF

// Inverter temperature (par 05.11, raw %)
IF _arrReadResults[7].quality = E_SignalQuality.Good THEN
	_telemetry.inverterTemp	:= UINT_TO_LREAL(_arrReadResults[7].valueUint);
END_IF

// Last fault code (par 04.11)
IF _arrReadResults[8].quality = E_SignalQuality.Good THEN
	_telemetry.faultCode	:= _arrReadResults[8].valueUint;
END_IF

// State label for HMI
IF _stsTripped THEN
	_stateString := 'Tripped';
ELSIF _arrReadResults[1].quality <> E_SignalQuality.Good THEN
	_stateString := 'No Comms';
ELSIF _stsSwOnInhibit THEN
	_stateString := 'Switch-On Inhibit';
ELSIF _stsRunning AND _stsAtSetpoint THEN
	_stateString := 'Running @ Setpoint';
ELSIF _stsRunning THEN
	_stateString := 'Running (Ramping)';
ELSIF _stsRdyOn THEN
	// RDY_RUN intentionally omitted: it is only asserted by the drive AFTER
	// OFF1 is released (CW bit 0 -> 1). RDY_ON with no inhibit is the real
	// "ready to be commanded" state.
	_stateString := 'Ready';
ELSE
	_stateString := 'Not Ready';
END_IF
END_METHOD

METHOD PRIVATE FaultHandler : BOOL
VAR_INPUT
END_VAR
// Each fault condition calls setFault separately with a unique description.
// The base class promotes the first one to the primary fault and emits any
// subsequent unique descriptions as 'Additional Fault - ...' warnings via
// the _extraFaults tracking. Combining descriptions into a single string
// would defeat that mechanism.

IF _stsTripped THEN
	setFault(1, CONCAT(CONCAT(CONCAT('Drive Fault: ', decodeFaultCode(_telemetry.faultCode)),
		' (code '), CONCAT(UINT_TO_STRING(_telemetry.faultCode), ')')));
END_IF

// Modbus driver exhausted reconnects (terminal)
IF _modbus.stsStatus.faulted THEN
	setFault(1, 'Modbus driver faulted (max reconnect attempts)');
END_IF

// No comms fault — fires whenever reads have been failing for >5s, regardless
// of driver state. Previously gated by currentState = Ready, which prevented
// the fault from firing during the very condition it was meant to catch.
IF _enabled AND _modbus.stsStatus.timeSinceLastGoodRead > T#5S THEN
	setFault(1, 'No Modbus comms');
END_IF

// Non-latching warnings
IF _stsAlarm THEN
	sendWarning(CONCAT(CONCAT(CONCAT('Drive alarm: ', decodeFaultCode(_telemetry.faultCode)),
		' (code '), CONCAT(UINT_TO_STRING(_telemetry.faultCode), ')')), 10);
END_IF

IF _enabled
   AND _arrReadResults[1].quality = E_SignalQuality.Good
   AND NOT _stsRemote THEN
	sendWarning('Drive in LOCAL mode (keypad)', 11);
END_IF

IF _stsSwOnInhibit AND _ctrlRunMode > 0 THEN
	sendWarning('Switch-on inhibit active; cannot start', 12);
END_IF
END_METHOD

METHOD PRIVATE decodeFaultCode : STRING
VAR_INPUT
	code : UINT;
END_VAR
// Common ACS580 fault codes. Not exhaustive — full list is in the ACS580
// firmware manual (3AUA0000078462). Add entries as you encounter them.
CASE code OF
	0:		decodeFaultCode := '';
	1080:	decodeFaultCode := 'Backup/restore timeout';
	2310:	decodeFaultCode := 'Overcurrent';
	2330:	decodeFaultCode := 'Earth leakage';
	2340:	decodeFaultCode := 'Short circuit';
	2381:	decodeFaultCode := 'IGBT overload';
	3130:	decodeFaultCode := 'Input phase loss';
	3181:	decodeFaultCode := 'Wiring or earth fault';
	3210:	decodeFaultCode := 'DC link overvoltage';
	3220:	decodeFaultCode := 'DC link undervoltage';
	3381:	decodeFaultCode := 'Output phase loss';
	4110:	decodeFaultCode := 'Control board overtemperature';
	4210:	decodeFaultCode := 'IGBT overtemperature';
	4290:	decodeFaultCode := 'Cooling';
	4310:	decodeFaultCode := 'Excess temperature';
	4380:	decodeFaultCode := 'Excess temperature difference';
	4981:	decodeFaultCode := 'External temperature 1';
	5080:	decodeFaultCode := 'Fan';
	5090:	decodeFaultCode := 'STO hardware failure';
	5091:	decodeFaultCode := 'Safe torque off';
	6481:	decodeFaultCode := 'Task overload';
	6487:	decodeFaultCode := 'Stack overflow';
	7081:	decodeFaultCode := 'Control panel loss';
	7082:	decodeFaultCode := 'Ext I/O comm loss';
	7121:	decodeFaultCode := 'Motor stall';
	7510:	decodeFaultCode := 'FBA A communication';
	7520:	decodeFaultCode := 'FBA B communication';
	7581:	decodeFaultCode := 'Drive-to-drive comm loss';
	9081:	decodeFaultCode := 'External event 1';
	9082:	decodeFaultCode := 'External event 2';
	9083:	decodeFaultCode := 'External event 3';
	9084:	decodeFaultCode := 'External event 4';
	9085:	decodeFaultCode := 'External event 5';
	20625:	decodeFaultCode := 'Safe torque off';			// 0x5091 hex - warning code
	36993:	decodeFaultCode := 'Safe torque off';			// 0x9081 hex - fault code
ELSE
	decodeFaultCode := 'Unknown fault';
END_CASE
END_METHOD

METHOD PRIVATE updateHMI : BOOL
VAR
END_VAR
HMI.HMIbaseDevice		:= HMIbaseDevice;
HMI.stsInterlocks		:= interlock.getHMIdata();

HMI.stsRunMode			:= _ctrlRunMode;
HMI.stsSetpoint			:= _ctrlSetpoint;

HMI.stsState			:= _stateString;
HMI.stsRunning			:= _stsRunning;
HMI.stsAtSetpoint		:= _stsAtSetpoint;
HMI.stsRemote			:= _stsRemote;
HMI.stsTripped			:= _stsTripped;
HMI.stsAlarm			:= _stsAlarm;

HMI.stsActualSpeed		:= _telemetry.actualSpeed;
HMI.stsMotorCurrent		:= _telemetry.motorCurrent;
HMI.stsDCBusVoltage		:= _telemetry.dcBusVoltage;
HMI.stsOutputFreq		:= _telemetry.outputFreq;
HMI.stsMotorTorque		:= _telemetry.motorTorque;
HMI.stsInverterTemp		:= _telemetry.inverterTemp;
HMI.stsFaultCode		:= stsFaultCode;
HMI.stsFaultText		:= stsFaultText;

HMI.stsCWRaw			:= _cwCurrent;
HMI.stsSWRaw			:= _swRaw;
HMI.stsCommsConnected	:= stsCommsConnected;
HMI.stsCommsFaulted		:= _modbus.stsStatus.faulted;
END_METHOD

METHOD FB_Init : BOOL
VAR_INPUT
	bInitRetains		: BOOL;	// TRUE: retain variables are initialized (reset warm / cold)
	bInCopyCode			: BOOL;	// TRUE: instance copied to copy code (online change)
	cfgDeviceName		: STRING;
	cfgEnable			: BOOL;
	cfgInitEventClass	: BOOL;
	cfgIPAddress		: STRING(15);
	cfgUnitID			: BYTE;
END_VAR
THIS^.cfgDeviceName		:= cfgDeviceName;
THIS^.cfgEnable			:= cfgEnable;
THIS^.cfgInitEventClass	:= cfgInitEventClass;
THIS^.cfgIPAddress		:= cfgIPAddress;
THIS^.cfgUnitID			:= cfgUnitID;
END_METHOD

END_FUNCTION_BLOCK

// ---- POUs/FBs/Devices/fb_Dev_VFD_DuraPulse.TcPOU
FUNCTION_BLOCK fb_Dev_VFD_DuraPulse EXTENDS abs_fb_Device
VAR_INPUT
	inpESTOPs_OK		: BOOL;		// 1 = ESTOPs healthy, 0 = ESTOP active
	inpMachineSTOP		: BOOL;
	inpCWAuxBitMask		: WORD;		// OR'd into outbound CW (0x2000) for app-specific bits
	inpExtFault			: BOOL;		// Trigger E.F. on the drive (0x2002 bit 0)
END_VAR

VAR PERSISTENT
	HMI					: ST_VFD_DuraPulse_HMI_Interface;
END_VAR

VAR
	_logSetpoint		: BOOL;
	// Embedded Modbus TCP client
	_modbus				: fb_Modbus_Driver;
	_modbusInit			: BOOL;

	// Read signal config. Two contiguous blocks reduce FC03 round-trips:
	//   - 0x2100..0x2106 (regs 1..7) cyclic status + primary telemetry
	//   - 0x210B..0x210C (regs 8..9) torque + rpm
	//   - 0x220E         (reg 10)    IGBT temperature
	_arrReadConfig		: ARRAY[1..10] OF ST_MBSignalConfig := [
		(modbusAddr := 48449, dataType := E_MBDataType.mbUInt16, tag := 'FaultWarn'),	// 0x2100
		(modbusAddr := 48450, dataType := E_MBDataType.mbUInt16, tag := 'SW'),			// 0x2101
		(modbusAddr := 48451, dataType := E_MBDataType.mbUInt16, tag := 'FCmdEcho'),	// 0x2102
		(modbusAddr := 48452, dataType := E_MBDataType.mbUInt16, tag := 'OutFreq'),		// 0x2103
		(modbusAddr := 48453, dataType := E_MBDataType.mbUInt16, tag := 'OutCurrent'),	// 0x2104
		(modbusAddr := 48454, dataType := E_MBDataType.mbUInt16, tag := 'DCBus'),		// 0x2105
		(modbusAddr := 48455, dataType := E_MBDataType.mbUInt16, tag := 'OutVoltage'),	// 0x2106
		(modbusAddr := 48460, dataType := E_MBDataType.mbInt16,  tag := 'Torque'),		// 0x210B
		(modbusAddr := 48461, dataType := E_MBDataType.mbInt16,  tag := 'MotorRPM'),	// 0x210C
		(modbusAddr := 48719, dataType := E_MBDataType.mbUInt16, tag := 'IGBTTemp')];	// 0x220E
	_arrReadResults		: ARRAY[1..10] OF ST_MBReadResult;

	// Write signal config: CW + Freq + bit-cmd (contiguous => single FC16)
	_arrWriteConfig		: ARRAY[1..3] OF ST_MBSignalConfig := [
		(modbusAddr := 48193, dataType := E_MBDataType.mbUInt16, tag := 'CW'),			// 0x2000
		(modbusAddr := 48194, dataType := E_MBDataType.mbUInt16, tag := 'FreqCmd'),		// 0x2001
		(modbusAddr := 48195, dataType := E_MBDataType.mbUInt16, tag := 'BitCmd')];		// 0x2002
	_arrWriteData		: ARRAY[1..3] OF ST_MBWriteData;

	// Application-level control signals
	_ctrlRunMode		: USINT;		// 0=stop, 1=fwd, 2=reverse
	_ctrlSetpoint		: LREAL;		// absolute Hz, 0..cfgMaxFreqHz
	_resetTrig			: R_TRIG;

	// Event-logging edge detection
	_lastLoggedRunMode	: USINT;
	_lastLoggedSetpoint	: LREAL;
	_trippedTrig		: R_TRIG;

	// CW state machine
	_cwState			: INT;			// 0=Idle, 1=Running, 2=FaultPending, 3=ResetSequence
	_cwCurrent			: WORD := 16#0001;	// init Stop (bits 1-0 = 01)
	_bitCmdCurrent		: WORD := 16#0000;	// 0x2002 bit commands (Reset, EF)
	_resetTimeout		: TON;
	_safetyStopActive	: BOOL;

	// Parsed status word
	_swRaw				: WORD;
	_stsRunBits			: BYTE;		// SW bits 0-1
	_stsDirBits			: BYTE;		// SW bits 3-4
	_stsJog				: BOOL;
	_stsFreqFromComm	: BOOL;		// SW bit 8
	_stsRemote			: BOOL;		// SW bit 10 — command via comm
	_stsParamsLocked	: BOOL;
	_stsRunning			: BOOL;		// SW bit 12
	_stsTripped			: BOOL;		// derived: low byte of 0x2100 != 0
	_stsAlarm			: BOOL;		// derived: high byte of 0x2100 != 0
	_stsDirection		: INT;		// +1 fwd, -1 rev, 0 stopped/transitioning

	// Engineering-unit telemetry
	_telemetry			: ST_VFD_DuraPulse_Telemetry;
	_stateString		: STRING;

	// Interlock array
	_interlocks			: ARRAY[1..10] OF BOOL;

	// Modbus configuration mirrors (set via cfg* properties before enable)
	_ipAddress			: STRING(15) := '192.168.1.50';
	_unitId				: BYTE := 1;
	_maxFreqHz			: LREAL := 60.0;	// must match drive P01.00
END_VAR

VAR_OUTPUT
	stsRunning			: BOOL;
	stsRemote			: BOOL;
	stsAlarm			: BOOL;
	stsTripped			: BOOL;
	stsDirection		: INT;		// +1 fwd, -1 rev, 0 stopped
	stsOutputFreq		: LREAL;	// Hz, signed
	stsMotorRPM			: LREAL;	// rpm, signed
	stsMotorCurrent		: LREAL;	// A
	stsDCBusVoltage		: LREAL;	// VDC
	stsOutputVoltage	: LREAL;	// VAC
	stsMotorTorque		: LREAL;	// %
	stsInverterTemp		: LREAL;	// degC
	stsFaultCode		: USINT;	// 0 unless drive is actively tripped
	stsFaultText		: STRING;
	stsWarningCode		: USINT;	// 0 unless warning active
	stsWarningText		: STRING;
	stsCommsConnected	: BOOL;
END_VAR

DeviceLogic();

// One-time Modbus driver configuration (properties lock after _initialized := TRUE)
IF NOT _modbusInit THEN
	_modbus.ipAddress				:= _ipAddress;
	_modbus.unitId					:= _unitId;
	_modbus.port					:= 502;
	_modbus.timeout					:= T#500MS;
	_modbus.pollInterval			:= T#50MS;
	_modbus.writeCycleInterval		:= T#100MS;
	_modbus.wordOrder				:= E_WordOrder.BigEndian;
	_modbus.maxConsecFails			:= 3;
	_modbus.reconnectDelay			:= T#2S;
	_modbus.maxReconnectAttempts	:= 10;
	_modbus.staleThreshold			:= T#2S;
	_modbus.readSignalCount			:= 10;
	_modbus.writeSignalCount		:= 3;
	_modbusInit := TRUE;
END_IF

// Drive the embedded Modbus client
_modbus(
	inpEnable			:= _enabled,
	inpPtrReadConfig	:= ADR(_arrReadConfig),
	inpPtrWriteConfig	:= ADR(_arrWriteConfig),
	inpPtrReadResults	:= ADR(_arrReadResults),
	inpPtrWriteData		:= ADR(_arrWriteData));
_modbus.cycle();

parseDriveFeedback();

// Interlocks
_interlocks[1] := inpESTOPs_OK;
cmdSetInterlock(1, 'ESTOPs OK', _interlocks[1]);

_interlocks[2] := NOT inpMachineSTOP;
cmdSetInterlock(2, 'Machine STOP Not Active', _interlocks[2]);

_interlocks[3] := _modbus.stsStatus.connected AND NOT _modbus.stsStatus.faulted;
cmdSetInterlock(3, 'Modbus comms OK', _interlocks[3]);

_interlocks[4] := _stsRemote;
cmdSetInterlock(4, 'Drive in Remote (comm) mode', _interlocks[4]);

_safetyStopActive := (NOT inpESTOPs_OK) OR inpMachineSTOP;

// HMI command surface — only honoured in manual mode
IF _enabled THEN
	IF NOT _inAuto THEN
		_ctrlRunMode	:= HMI.ocmdRunMode;
		_ctrlSetpoint	:= HMI.ocmdSetpoint;
	END_IF
END_IF

_resetTrig(CLK := HMI.ocmdReset);
IF _resetTrig.Q THEN
	cmdReset();
END_IF

FaultHandler();

// Interlock enforcement
IF NOT interlock.outInterlockOK THEN
	_ctrlRunMode	:= 0;
	HMI.ocmdRunMode	:= 0;
END_IF

controlWordSequencer();

// Marshal CW + freq + bit-cmd into Modbus write buffers
_arrWriteData[1].valueUint	:= WORD_TO_UINT(_cwCurrent OR inpCWAuxBitMask);
_arrWriteData[2].valueUint	:= LREAL_TO_UINT(LIMIT(0.0, _ctrlSetpoint, _maxFreqHz) * 100.0);
// 0x2002 bit 0 = E.F. trigger (pulse from caller), bit 1 = reset (managed by sequencer)
_arrWriteData[3].valueUint	:= WORD_TO_UINT(_bitCmdCurrent OR BOOL_TO_WORD(inpExtFault));

// Event-based logging
IF _ctrlRunMode <> _lastLoggedRunMode THEN
	CASE _ctrlRunMode OF
		0:	sendLog('Stop command', 1);
		1:	sendLog(CONCAT(CONCAT('Run forward @ ', LREAL_TO_STRING(_ctrlSetpoint)), ' Hz'), 1);
		2:	sendLog(CONCAT(CONCAT('Run reverse @ ', LREAL_TO_STRING(_ctrlSetpoint)), ' Hz'), 1);
	END_CASE
	_lastLoggedRunMode := _ctrlRunMode;
END_IF

IF ABS(_ctrlSetpoint - _lastLoggedSetpoint) >= 0.1 THEN
	IF _logSetpoint THEN
		sendLog(CONCAT(CONCAT('Setpoint = ', LREAL_TO_STRING(_ctrlSetpoint)), ' Hz'), 2);
		_lastLoggedSetpoint := _ctrlSetpoint;
	END_IF
END_IF

_trippedTrig(CLK := _stsTripped);
IF _trippedTrig.Q THEN
	sendLog(CONCAT('Drive tripped, fault code ', USINT_TO_STRING(_telemetry.faultCode)), 3);
END_IF

updateHMI();

// Public outputs
stsRunning			:= _stsRunning;
stsRemote			:= _stsRemote;
stsAlarm			:= _stsAlarm;
stsTripped			:= _stsTripped;
stsDirection		:= _stsDirection;
stsOutputFreq		:= _telemetry.outputFreq;
stsMotorRPM			:= _telemetry.motorRPM;
stsMotorCurrent		:= _telemetry.motorCurrent;
stsDCBusVoltage		:= _telemetry.dcBusVoltage;
stsOutputVoltage	:= _telemetry.outputVoltage;
stsMotorTorque		:= _telemetry.motorTorque;
stsInverterTemp		:= _telemetry.inverterTemp;
// Gate fault/warning text by active condition. The drive does not latch
// these codes once the condition clears, but we still want explicit text
// suppression on the operator-facing outputs.
IF _stsTripped THEN
	stsFaultCode	:= _telemetry.faultCode;
	stsFaultText	:= decodeAlarmCode(_telemetry.faultCode);
ELSE
	stsFaultCode	:= 0;
	stsFaultText	:= '';
END_IF
IF _stsAlarm THEN
	stsWarningCode	:= _telemetry.warningCode;
	stsWarningText	:= decodeAlarmCode(_telemetry.warningCode);
ELSE
	stsWarningCode	:= 0;
	stsWarningText	:= '';
END_IF
// AND with signal quality so this agrees with the 'No Comms' state string.
// Driver's connected flag lags reality (only drops after maxConsecFails);
// signal quality flips on the first failed read.
stsCommsConnected	:= _modbus.stsStatus.connected AND (_arrReadResults[2].quality = E_SignalQuality.Good);

PROPERTY cfgIPAddress : STRING(15)
GET
cfgIPAddress := _ipAddress;
END_GET
SET
_ipAddress := cfgIPAddress;
END_SET
END_PROPERTY

PROPERTY cfgLogSetpoint : BOOL
GET
cfgLogSetpoint := _logSetpoint;
END_GET
SET
_logsetpoint := cfgLogSetpoint;
END_SET
END_PROPERTY

// Drive-side maximum frequency (P01.00). Used to clamp setpoint client-side.
PROPERTY cfgMaxFreqHz : LREAL
GET
cfgMaxFreqHz := _maxFreqHz;
END_GET
SET
IF cfgMaxFreqHz > 0.0 THEN
	_maxFreqHz := cfgMaxFreqHz;
END_IF
END_SET
END_PROPERTY

PROPERTY cfgUnitID : BYTE
GET
cfgUnitID := _unitId;
END_GET
SET
_unitId := cfgUnitID;
END_SET
END_PROPERTY

METHOD PUBLIC cmdEnable : BOOL
VAR_INPUT
	command		: USINT;	// 0=stop, 1=run forward, 2=run reverse
END_VAR
IF command <= 2 THEN
	_ctrlRunMode := command;
END_IF
END_METHOD

METHOD PUBLIC cmdReset : BOOL
setFault(0, '');
IF _stsTripped THEN
	_cwState := 3;
END_IF
// A driver that gave up after maxReconnectAttempts restarts on reset (it no longer needs a
// PLC restart to recover).
IF _modbus.stsStatus.faulted THEN
	_modbus.cmdReset();
END_IF
END_METHOD

METHOD PUBLIC cmdSetpoint : BOOL
VAR_INPUT
	setpoint	: LREAL;	// absolute Hz, 0..cfgMaxFreqHz
END_VAR
_ctrlSetpoint := LIMIT(0.0, setpoint, _maxFreqHz);
END_METHOD

METHOD PRIVATE controlWordSequencer : BOOL
VAR_INPUT
END_VAR
// DuraPulse CW values (register 0x2000):
//   0x0001 = Stop (bits 1-0 = 01)
//   0x0012 = Run forward (run + FWD)
//   0x0022 = Run reverse (run + REV)
//
// Reset is performed via 0x2002 bit 1 (separate register), pulsed by state 3.
// The drive does not require an ABB-style "ready" precondition — it will
// accept Run directly from Stop once any fault is cleared.

// Default to no bit commands (reset bit clears outside state 3)
_bitCmdCurrent := 16#0000;

CASE _cwState OF
	0:	// Idle / Stopped
		_cwCurrent := 16#0001;
		IF _ctrlRunMode > 0
		   AND NOT _stsTripped
		   AND NOT _safetyStopActive THEN
			_cwState := 1;
		ELSIF _stsTripped THEN
			_cwState := 2;
		END_IF

	1:	// Running
		IF _stsTripped THEN
			_cwState := 2;
		ELSIF _ctrlRunMode = 0 OR _safetyStopActive THEN
			_cwState := 0;
		ELSIF _ctrlRunMode = 1 THEN
			_cwCurrent := 16#0012;		// run forward
		ELSIF _ctrlRunMode = 2 THEN
			_cwCurrent := 16#0022;		// run reverse
		END_IF

	2:	// FaultPending — wait for reset
		_cwCurrent := 16#0001;
		IF NOT _stsTripped THEN
			_cwState := 0;
		END_IF

	3:	// ResetSequence — hold reset bit until fault clears (max 3s)
		_cwCurrent := 16#0001;
		_bitCmdCurrent := 16#0002;		// 0x2002 bit 1 = reset
		_resetTimeout(IN := TRUE, PT := T#3S);
		IF NOT _stsTripped THEN
			_cwState := 0;
			_resetTimeout(IN := FALSE);
		ELSIF _resetTimeout.Q THEN
			setFault(1, 'Fault reset did not clear after 3s');
			_cwState := 2;
			_resetTimeout(IN := FALSE);
		END_IF
END_CASE
END_METHOD

METHOD PRIVATE decodeAlarmCode : STRING
VAR_INPUT
	code : USINT;
END_VAR
// Common GS20(X) / Delta MS300 fault & warning codes. Not exhaustive — full
// list is in GS20 manual Chapter 6 (Maintenance and Troubleshooting).
// Both fault (low byte of 0x2100) and warning (high byte) use the same
// numbering scheme, so one decode function covers both.
CASE code OF
	0:		decodeAlarmCode := '';
	1:		decodeAlarmCode := 'Overcurrent during acceleration (ocA)';
	2:		decodeAlarmCode := 'Overcurrent during deceleration (ocd)';
	3:		decodeAlarmCode := 'Overcurrent during steady state (ocn)';
	4:		decodeAlarmCode := 'Ground fault (GFF)';
	5:		decodeAlarmCode := 'IGBT short circuit (occ)';
	6:		decodeAlarmCode := 'Overcurrent at stop (ocS)';
	7:		decodeAlarmCode := 'Overvoltage during acceleration (ovA)';
	8:		decodeAlarmCode := 'Overvoltage during deceleration (ovd)';
	9:		decodeAlarmCode := 'Overvoltage during steady state (ovn)';
	10:		decodeAlarmCode := 'Overvoltage at stop (ovS)';
	11:		decodeAlarmCode := 'Low voltage during acceleration (LvA)';
	12:		decodeAlarmCode := 'Low voltage during deceleration (Lvd)';
	13:		decodeAlarmCode := 'Low voltage during steady state (Lvn)';
	14:		decodeAlarmCode := 'Low voltage at stop (LvS)';
	15:		decodeAlarmCode := 'Phase loss protection (OrP)';
	16:		decodeAlarmCode := 'IGBT overheat (oH1)';
	17:		decodeAlarmCode := 'Capacitor overheat (oH2)';
	18:		decodeAlarmCode := 'IGBT temperature sensor error (tH1o)';
	19:		decodeAlarmCode := 'Capacitor temperature sensor error (tH2o)';
	21:		decodeAlarmCode := 'Drive overload (oL)';
	22:		decodeAlarmCode := 'Electronic thermal relay 1 (EoL1)';
	23:		decodeAlarmCode := 'Electronic thermal relay 2 (EoL2)';
	24:		decodeAlarmCode := 'Motor PTC overheat (oH3)';
	26:		decodeAlarmCode := 'Over-torque 1 (ot1)';
	27:		decodeAlarmCode := 'Over-torque 2 (ot2)';
	28:		decodeAlarmCode := 'Low current (uC)';
	31:		decodeAlarmCode := 'EEPROM read error (cF2)';
	33:		decodeAlarmCode := 'U-phase current detection error (cd1)';
	34:		decodeAlarmCode := 'V-phase current detection error (cd2)';
	35:		decodeAlarmCode := 'W-phase current detection error (cd3)';
	36:		decodeAlarmCode := 'Clamp current detection error (Hd0)';
	37:		decodeAlarmCode := 'Over-current detection error (Hd1)';
	40:		decodeAlarmCode := 'Auto-tuning error (AUE)';
	41:		decodeAlarmCode := 'PID feedback loss (AFE)';
	48:		decodeAlarmCode := 'Analog current input loss (ACE)';
	49:		decodeAlarmCode := 'External fault input (EF)';
	50:		decodeAlarmCode := 'Emergency stop (EF1)';
	51:		decodeAlarmCode := 'External base block (bb)';
	52:		decodeAlarmCode := 'Password fault (Pcod)';
	54:		decodeAlarmCode := 'Communication error (CE1)';
	55:		decodeAlarmCode := 'Communication error (CE2)';
	56:		decodeAlarmCode := 'Communication error (CE3)';
	57:		decodeAlarmCode := 'Communication error (CE4)';
	58:		decodeAlarmCode := 'Modbus comm time-out (CE10)';
	60:		decodeAlarmCode := 'Brake transistor error (bF)';
	61:		decodeAlarmCode := 'Y-connection / delta-connection switch error (ydc)';
	62:		decodeAlarmCode := 'Deceleration energy backup error (dEb)';
	72:		decodeAlarmCode := 'STO loss 1 (STL1)';
	76:		decodeAlarmCode := 'Safe torque off (STo)';
	77:		decodeAlarmCode := 'STO loss 2 (STL2)';
	78:		decodeAlarmCode := 'STO loss 3 (STL3)';
	79:		decodeAlarmCode := 'U-phase output phase loss (OPHL)';
	80:		decodeAlarmCode := 'V-phase output phase loss (OPHL)';
	81:		decodeAlarmCode := 'W-phase output phase loss (OPHL)';
	82:		decodeAlarmCode := 'Output phase loss (OPHL)';
	87:		decodeAlarmCode := 'Drive overload (oL3)';
	101:	decodeAlarmCode := 'CANopen software disconnect 1 (CGdE)';
	121:	decodeAlarmCode := 'Internal communication error (CP20)';
ELSE
	decodeAlarmCode := 'Unknown code';
END_CASE
END_METHOD

METHOD PRIVATE FaultHandler : BOOL
VAR_INPUT
END_VAR
// Each fault condition calls setFault separately so the base class can
// promote the first one to the primary fault and report subsequent ones
// as 'Additional Fault - ...' warnings.

IF _stsTripped THEN
	setFault(1, CONCAT(CONCAT(CONCAT('Drive Fault: ', decodeAlarmCode(_telemetry.faultCode)),
		' (code '), CONCAT(USINT_TO_STRING(_telemetry.faultCode), ')')));
END_IF

// Modbus driver exhausted reconnects (terminal)
IF _modbus.stsStatus.faulted THEN
	setFault(1, 'Modbus driver faulted (max reconnect attempts)');
END_IF

// No comms fault — fires whenever reads have been failing for >5s
IF _enabled AND _modbus.stsStatus.timeSinceLastGoodRead > T#5S THEN
	setFault(1, 'No Modbus comms');
END_IF

// Non-latching warnings
IF _stsAlarm THEN
	sendWarning(CONCAT(CONCAT(CONCAT('Drive warning: ', decodeAlarmCode(_telemetry.warningCode)),
		' (code '), CONCAT(USINT_TO_STRING(_telemetry.warningCode), ')')), 10);
END_IF

IF _enabled
   AND _arrReadResults[2].quality = E_SignalQuality.Good
   AND NOT _stsRemote THEN
	sendWarning('Drive command source is not Communication (local/keypad)', 11);
END_IF
END_METHOD

METHOD FB_Init : BOOL
VAR_INPUT
	bInitRetains		: BOOL;	// TRUE: retain variables are initialized (reset warm / cold)
	bInCopyCode			: BOOL;	// TRUE: instance copied to copy code (online change)
	cfgDeviceName		: STRING;
	cfgEnable			: BOOL;
	cfgInitEventClass	: BOOL;
	cfgIPAddress		: STRING(15);
	cfgUnitID			: BYTE;
	cfgMaxFreqHz		: LREAL;
END_VAR
THIS^.cfgDeviceName		:= cfgDeviceName;
THIS^.cfgEnable			:= cfgEnable;
THIS^.cfgInitEventClass	:= cfgInitEventClass;
THIS^.cfgIPAddress		:= cfgIPAddress;
THIS^.cfgUnitID			:= cfgUnitID;
IF cfgMaxFreqHz > 0.0 THEN
	THIS^.cfgMaxFreqHz	:= cfgMaxFreqHz;
END_IF
END_METHOD

METHOD PRIVATE parseDriveFeedback : BOOL
VAR
	_faultWarn	: WORD;
END_VAR
// 0x2100: low byte = fault, high byte = warning
IF _arrReadResults[1].quality = E_SignalQuality.Good THEN
	_faultWarn				:= UINT_TO_WORD(_arrReadResults[1].valueUint);
	_telemetry.faultCode	:= WORD_TO_USINT(_faultWarn AND 16#00FF);
	_telemetry.warningCode	:= WORD_TO_USINT(SHR(_faultWarn AND 16#FF00, 8));
	_stsTripped				:= _telemetry.faultCode <> 0;
	_stsAlarm				:= _telemetry.warningCode <> 0;
END_IF

// 0x2101: status word
IF _arrReadResults[2].quality = E_SignalQuality.Good THEN
	_swRaw				:= UINT_TO_WORD(_arrReadResults[2].valueUint);
	_stsRunBits			:= WORD_TO_BYTE(_swRaw AND 16#0003);				// bits 0-1
	_stsJog				:= (_swRaw AND 16#0004) <> 0;						// bit 2
	_stsDirBits			:= WORD_TO_BYTE(SHR(_swRaw AND 16#0018, 3));		// bits 3-4
	_stsFreqFromComm	:= (_swRaw AND 16#0100) <> 0;						// bit 8
	_stsRemote			:= (_swRaw AND 16#0400) <> 0;						// bit 10
	_stsParamsLocked	:= (_swRaw AND 16#0800) <> 0;						// bit 11
	_stsRunning			:= (_swRaw AND 16#1000) <> 0;						// bit 12

	// Direction (0=fwd, 3=rev, 1/2=transition)
	CASE _stsDirBits OF
		0:	_stsDirection := SEL(_stsRunning, 0, 1);	// fwd only meaningful while running
		3:	_stsDirection := -1;
	ELSE
		_stsDirection := 0;		// transitioning
	END_CASE
END_IF

// 0x2103: output frequency (UInt, 0.01 Hz). Sign from direction.
IF _arrReadResults[4].quality = E_SignalQuality.Good THEN
	_telemetry.outputFreq	:= UINT_TO_LREAL(_arrReadResults[4].valueUint) / 100.0;
	IF _stsDirection < 0 THEN
		_telemetry.outputFreq := -_telemetry.outputFreq;
	END_IF
END_IF

// 0x2104: output current (0.01 A)
IF _arrReadResults[5].quality = E_SignalQuality.Good THEN
	_telemetry.motorCurrent	:= UINT_TO_LREAL(_arrReadResults[5].valueUint) / 100.0;
END_IF

// 0x2105: DC bus voltage (0.1 VDC)
IF _arrReadResults[6].quality = E_SignalQuality.Good THEN
	_telemetry.dcBusVoltage	:= UINT_TO_LREAL(_arrReadResults[6].valueUint) / 10.0;
END_IF

// 0x2106: output voltage (0.1 VAC)
IF _arrReadResults[7].quality = E_SignalQuality.Good THEN
	_telemetry.outputVoltage := UINT_TO_LREAL(_arrReadResults[7].valueUint) / 10.0;
END_IF

// 0x210B: output torque (signed 0.1 %)
IF _arrReadResults[8].quality = E_SignalQuality.Good THEN
	_telemetry.motorTorque	:= INT_TO_LREAL(_arrReadResults[8].valueInt) / 10.0;
END_IF

// 0x210C: actual motor speed (signed rpm)
IF _arrReadResults[9].quality = E_SignalQuality.Good THEN
	_telemetry.motorRPM		:= INT_TO_LREAL(_arrReadResults[9].valueInt);
END_IF

// 0x220E: IGBT temperature (0.1 degC)
IF _arrReadResults[10].quality = E_SignalQuality.Good THEN
	_telemetry.inverterTemp	:= UINT_TO_LREAL(_arrReadResults[10].valueUint) / 10.0;
END_IF

// State label for HMI
IF _stsTripped THEN
	_stateString := 'Tripped';
ELSIF _arrReadResults[2].quality <> E_SignalQuality.Good THEN
	_stateString := 'No Comms';
ELSIF NOT _stsRemote THEN
	_stateString := 'Local Mode';
ELSIF _stsRunBits = 2#11 THEN
	_stateString := 'Running';
ELSIF _stsRunBits = 2#10 THEN
	_stateString := 'Standby';
ELSIF _stsRunBits = 2#01 THEN
	_stateString := 'Decelerating';
ELSE
	_stateString := 'Stopped';
END_IF
END_METHOD

METHOD PRIVATE updateHMI : BOOL
VAR
END_VAR
HMI.HMIbaseDevice		:= HMIbaseDevice;
HMI.stsInterlocks		:= interlock.getHMIdata();

HMI.stsRunMode			:= _ctrlRunMode;
HMI.stsSetpoint			:= _ctrlSetpoint;

HMI.stsState			:= _stateString;
HMI.stsRunning			:= _stsRunning;
HMI.stsRemote			:= _stsRemote;
HMI.stsTripped			:= _stsTripped;
HMI.stsAlarm			:= _stsAlarm;
HMI.stsDirection		:= _stsDirection;

HMI.stsOutputFreq		:= _telemetry.outputFreq;
HMI.stsMotorRPM			:= _telemetry.motorRPM;
HMI.stsMotorCurrent		:= _telemetry.motorCurrent;
HMI.stsDCBusVoltage		:= _telemetry.dcBusVoltage;
HMI.stsOutputVoltage	:= _telemetry.outputVoltage;
HMI.stsMotorTorque		:= _telemetry.motorTorque;
HMI.stsInverterTemp		:= _telemetry.inverterTemp;
HMI.stsFaultCode		:= stsFaultCode;
HMI.stsFaultText		:= stsFaultText;
HMI.stsWarningCode		:= stsWarningCode;
HMI.stsWarningText		:= stsWarningText;

HMI.stsCWRaw			:= _cwCurrent;
HMI.stsSWRaw			:= _swRaw;
HMI.stsCommsConnected	:= stsCommsConnected;
HMI.stsCommsFaulted		:= _modbus.stsStatus.faulted;
END_METHOD

END_FUNCTION_BLOCK

// ---- POUs/FBs/Devices/fb_Dev_WebRelay.TcPOU
FUNCTION_BLOCK fb_Dev_WebRelay EXTENDS abs_fb_Device

VAR_INPUT
	inpRelayCmd	: BOOL;
END_VAR

VAR
	_commFault				: BOOL;
	_modbus_IF				: ST_Modbus_Commands;
	_modbus_cfg				: ST_Modbus_Device_Config;
	_modbus_WC_state		: INT;
	_modbus_RC_state		: INT;
	_DIReadDelay			: TON;
	_DIReadDelayTrig		: BOOL;
	_DIState				: BOOL;
	_DOWriteDelay			: TON;
	_DOWriteDelayTrig		: BOOL;
	_setDO					: BOOL;

END_VAR

VAR_OUTPUT
	stsDI	: BOOL;
	stsDO	: BOOL;
END_VAR

DeviceLogic();
Interlock.name := _DeviceName;
Interlock(inpConfig := _dataInterlock);

//Set device config for WriteSingleCoil
_modbus_IF.WriteSingleCoil.sIPAddr 		:= _modbus_cfg.cfgIP_address;
_modbus_IF.WriteSingleCoil.nTCPPort 	:= _modbus_cfg.cfgTCPPort;
_modbus_IF.WriteSingleCoil.nUnitID		:= _modbus_cfg.cfgUnitID;
_modbus_IF.WriteSingleCoil.tTimeout 	:= _modbus_cfg.cfgTimeout;
_modbus_IF.WriteSingleCoil.nMBAddr		:= 1;

_modbus_IF.ReadInputs.sIPAddr			:= _modbus_cfg.cfgIP_address;
_modbus_IF.ReadInputs.nTCPPort			:= _modbus_cfg.cfgTCPPort;
_modbus_IF.ReadInputs.nUnitID			:= _modbus_cfg.cfgUnitID;
_modbus_IF.ReadInputs.tTimeout			:= _modbus_cfg.cfgTimeout;
_modbus_IF.ReadInputs.nMBAddr			:= 0;

_DIReadDelay(IN:=_DIReadDelayTrig, PT:=T#250MS);
_DOWriteDelay(IN:=_DOWriteDelayTrig, PT:=T#250MS);
_modbus_IF.ReadInputs();
_modbus_IF.WriteSingleCoil();

// Read the DI alue
cmdReadDI();

FaultHandler();

// Set the relay based on fb input unless it's faulted
IF NOT stsFaulted THEN
	_setDO := inpRelayCmd;
ELSE
	_setDO := FALSE;
END_IF

cmdSetDO(_setDO);

stsDI := _DIState;
stsDO := _setDO;

PROPERTY cfgDeviceName : string
GET
cfgDeviceName := _devicename;
END_GET
SET
_devicename := cfgDeviceName;
END_SET
END_PROPERTY

PROPERTY cfgEnable : bool
GET
cfgEnable := _enabled;
END_GET
SET
_enabled := cfgEnable;
END_SET
END_PROPERTY

PROPERTY cfgModbusConfig : ST_Modbus_Device_Config
GET
cfgModbusConfig := _modbus_cfg;
END_GET
SET
_modbus_cfg := cfgModbusConfig;
END_SET
END_PROPERTY

METHOD cmdReadDI : BOOL
VAR_INPUT
END_VAR
CASE _modbus_RC_state OF
	0:
		_modbus_IF.ReadInputs.nQuantity := SIZEOF(_DIState);
		_modbus_IF.ReadInputs.cbLength  := SIZEOF(_DIState);
		_modbus_IF.ReadInputs.pDestAddr := ADR(_DIState);
		_modbus_IF.ReadInputs.bExecute  := TRUE;
		_modbus_RC_state := 1;
	1:
		_modbus_IF.ReadInputs.bExecute := FALSE;
		_DIReadDelayTrig := TRUE;
		IF _DIReadDelay.Q THEN
			_DIReadDelayTrig := FALSE;
			_modbus_RC_state := 0;
		END_IF
END_CASE
END_METHOD

METHOD cmdReset : BOOL
IF stsFaulted THEN
	setFault(0,'');
	IF _commFault = TRUE THEN
		_commFault := FALSE;
		_modbus_IF.WriteSingleCoil.bExecute:= FALSE;
		_modbus_WC_state  := 0;
	END_IF
END_IF
END_METHOD

METHOD PUBLIC cmdSetDO : BOOL
VAR_INPUT
	setRequest	: Bool;
END_VAR
CASE _modbus_WC_state OF
	0:
		IF setRequest = TRUE THEN
			_modbus_IF.WriteSingleCoil.nValue := 65280;
		ELSE
			_modbus_IF.WriteSingleCoil.nValue := 0;
		END_IF
		
		_modbus_IF.WriteSingleCoil.bExecute := TRUE;
		IF _modbus_IF.WriteSingleCoil.bBusy = TRUE THEN
			_modbus_WC_state := 1;
		END_IF
	1:
		_modbus_IF.WriteSingleCoil.bExecute := FALSE;
		_DOWriteDelayTrig := TRUE;
		IF _DOWriteDelay.Q THEN
			_DOWriteDelayTrig := FALSE;
			_modbus_WC_state := 0;
		END_IF
END_CASE
END_METHOD

METHOD FaultHandler : BOOL
VAR_INPUT
END_VAR
IF _modbus_IF.WriteSingleCoil.bError THEN
	setFault(1,'Comms. Write Fault');
	_commFault := TRUE;
END_IF

IF _modbus_IF.ReadInputs.bError THEN
	setFault(1,'Comms. Read Fault');
	_commFault := TRUE;
END_IF

IF NOT interlock.outInterlockOK THEN
	setFault(1,CONCAT('I_NOK - ',Interlock.stsFirstOut));
END_IF
END_METHOD

//FB_Init is always available implicitly and it is used primarily for initialization.
//The return value is not evaluated. For a specific influence, you can also declare the
//methods explicitly and provide additional code there with the standard initialization
//code. You can evaluate the return value.
METHOD FB_Init: BOOL
VAR_INPUT
    bInitRetains		: BOOL; // TRUE: the retain variables are initialized (reset warm / reset cold)
    bInCopyCode			: BOOL;  // TRUE: the instance will be copied to the copy code afterward (online change)  
	cfgDeviceName		: STRING;
	cfgEnable			: BOOL; 
	cfgInitEventClass	: BOOL;    
END_VAR
THIS^.cfgDeviceName 		:= 		cfgDeviceName; 		
THIS^.cfgEnable 			:= 	    cfgEnable;
THIS^.cfgInitEventClass		:= 		cfgInitEventClass;
END_METHOD

END_FUNCTION_BLOCK

// ---- POUs/FBs/Devices/fb_Dev_ControlValve_Modulating_REAL.TcPOU
FUNCTION_BLOCK fb_Dev_ControlValve_Modulating_REAL
VAR_INPUT
	IO_valveFeedback	: LREAL;
	IO_valveOutput		: POINTER TO REAL;
	inpAuto				: BOOL;
	inpReset			: BOOL;
	inpInterlockBypass	: BOOL;
	faultMonitor		: POINTER TO fb_FaultMonitor;
END_VAR

VAR
	valveFeedback_scaled	: LREAL;
	_valveName				: STRING;
	Valve					: fb_Dev_ControlValve_Modulating(cfgDeviceName := _valveName, cfgEnable := TRUE, cfgInitEventClass := TRUE);
	_valvePositionCmd		: LREAL;
	
END_VAR
VAR_OUTPUT
	outValvePosition	: LREAL;
	stsValveFeedback	: LREAL;
END_VAR

//INPUTS AND OUTPUTS FOR THIS FB VARIANT ARE SCALED ANALOG VALUES IN VOLTS
valveFeedback_scaled := F_AnalogToEngUnit(IO_valveFeedback, 2, 10, 0, 100);

Valve(inpAuto := inpAuto, inpReset := inpReset, inpInterlockBypass := inpInterlockBypass, faultMonitor:=faultMonitor
		, inpValvePosition := valveFeedback_scaled);
		
outValvePosition := Valve.outValvePosition;
stsValveFeedback := Valve.stsValveFeedback;

Valve.valvePosition := _valvePositionCmd;

		
IO_valveOutput^ := F_AnalogToEngUnit(TO_LREAL(Valve.outValvePosition), 0, 100, 2, 10);

PROPERTY cmdSetValvePosition : LREAL
SET
_valvePositionCmd := cmdSetValvePosition;
END_SET
END_PROPERTY

//FB_Init is always available implicitly and it is used primarily for initialization.
//The return value is not evaluated. For a specific influence, you can also declare the
//methods explicitly and provide additional code there with the standard initialization
//code. You can evaluate the return value.
METHOD FB_Init: BOOL
VAR_INPUT
    bInitRetains: BOOL; // TRUE: the retain variables are initialized (reset warm / reset cold)
    bInCopyCode: BOOL;  // TRUE: the instance will be copied to the copy code afterward (online change) 
	cfgDeviceName	: STRING;  
END_VAR
THIS^._valveName 			:= cfgDeviceName;
THIS^.Valve.cfgDeviceName 	:= cfgDeviceName;
END_METHOD

END_FUNCTION_BLOCK

// ---- POUs/FBs/Devices/fb_Dev_IsolationMonitor.TcPOU
FUNCTION_BLOCK fb_Dev_IsolationMonitor EXTENDS abs_fb_device

VAR_INPUT
	IO_IN_DeviceTrip	: POINTER TO BOOL;
	IO_IN_DeviceWarning	: POINTER TO BOOL;
	IO_OUT_TripReset	: POINTER TO BOOL;
	IO_OUT_Test			: POINTER TO BOOL;
END_VAR

VAR
	_modbus_IF				: ST_Modbus_Commands;
	_modbus_cfg				: ST_Modbus_Device_Config;
	_RegReadTimer			: TON;
	_RegWriteTimer			: TON;
	_RegReadState			:INT := 0;
	_RegRead				: ARRAY [1..84] OF BYTE;
	_IsoMon_DeviceSignals	: ST_IsoMon_MBIF;
	HMI						: ST_IsoMon_HMI_Interface;
	HMI_DeviceSignals		: ST_IsoMon_DeviceSignals;
	TOFReset				: TOF;
	TOFResetTrig			: BOOL;
	TOFTest					: TOF;
	TOFTestTrig				: BOOL;
	_cmdResetTrip			: BOOL;
	_commOK					: BOOL;		// TRUE after the last register read succeeded

	
END_VAR

VAR_OUTPUT
	stsInsulationResistance	: REAL;
	stsCommOK				: BOOL;		// FALSE = the readings below are NOT current (read failed or not yet read)
END_VAR

DeviceLogic();
Interlock.name := _DeviceName;
Interlock(inpConfig := _dataInterlock);

FaultHandler();

//Set device config for Modbus interface
_modbus_IF.ReadRegisters.sIPAddr	:= _modbus_cfg.cfgIP_address;
_modbus_IF.ReadRegisters.nTCPPort 	:= _modbus_cfg.cfgTCPPort;
_modbus_IF.ReadRegisters.nUnitID	:= _modbus_cfg.cfgUnitID;
_modbus_IF.ReadRegisters.tTimeout 	:= _modbus_cfg.cfgTimeout;

IF _enabled THEN	
	_modbus_IF.ReadRegisters();
END_IF

//Read Registers (parsed only when a read completes without error - see cmdReadRegisters)
IF _enabled THEN
	cmdReadRegisters();
ELSE
	_commOK := FALSE;
END_IF
stsCommOK := _commOK;

_RegReadTimer(IN := NOT _RegReadTimer.Q, PT := T#0.1S);
IF _RegReadTimer.Q THEN
	IF _RegReadState = 900 THEN
		_RegReadState := 0;
	END_IF
END_IF

TOFReset(IN:=TOFResetTrig, PT:= T#1S);
TOFTest(IN:=TOFTestTrig, PT:= T#1S);

//DataTask.IsoMon_InsulationResistance	:= _IsoMon_DeviceSignals.insulationResistance.value / 1000;

updateHMI();

stsInsulationResistance := HMI_deviceSignals.insulationResistance_kOhm;

PROPERTY cfgModbusConfig : ST_Modbus_Device_Config
GET
cfgModbusConfig := _modbus_cfg;
END_GET
SET
_modbus_cfg := cfgModbusConfig;
END_SET
END_PROPERTY

METHOD PRIVATE cmdParseRegisters : BOOL
VAR_INPUT
END_VAR
// 0x2000: insulationResistance
_IsoMon_DeviceSignals.insulationResistance.bytes[1] := _RegRead[3];
_IsoMon_DeviceSignals.insulationResistance.bytes[2] := _RegRead[4];
_IsoMon_DeviceSignals.insulationResistance.bytes[3] := _RegRead[1];
_IsoMon_DeviceSignals.insulationResistance.bytes[4] := _RegRead[2];

// 0x2002: minInsulationValue
_IsoMon_DeviceSignals.minInsulationValue.bytes[1] := _RegRead[7];
_IsoMon_DeviceSignals.minInsulationValue.bytes[2] := _RegRead[8];
_IsoMon_DeviceSignals.minInsulationValue.bytes[3] := _RegRead[5];
_IsoMon_DeviceSignals.minInsulationValue.bytes[4] := _RegRead[6];

// 0x2004: systemLeakageCapacitance
_IsoMon_DeviceSignals.systemLeakageCapacitance.bytes[1] := _RegRead[11];
_IsoMon_DeviceSignals.systemLeakageCapacitance.bytes[2] := _RegRead[12];
_IsoMon_DeviceSignals.systemLeakageCapacitance.bytes[3] := _RegRead[9];
_IsoMon_DeviceSignals.systemLeakageCapacitance.bytes[4] := _RegRead[10];

// 0x2006: voltageL1L2
_IsoMon_DeviceSignals.voltageL1L2.bytes[1] := _RegRead[15];
_IsoMon_DeviceSignals.voltageL1L2.bytes[2] := _RegRead[16];
_IsoMon_DeviceSignals.voltageL1L2.bytes[3] := _RegRead[13];
_IsoMon_DeviceSignals.voltageL1L2.bytes[4] := _RegRead[14];

// 0x2008: voltageL1L3
_IsoMon_DeviceSignals.voltageL1L3.bytes[1] := _RegRead[19];
_IsoMon_DeviceSignals.voltageL1L3.bytes[2] := _RegRead[20];
_IsoMon_DeviceSignals.voltageL1L3.bytes[3] := _RegRead[17];
_IsoMon_DeviceSignals.voltageL1L3.bytes[4] := _RegRead[18];

// 0x200A: voltageL2L3
_IsoMon_DeviceSignals.voltageL2L3.bytes[1] := _RegRead[23];
_IsoMon_DeviceSignals.voltageL2L3.bytes[2] := _RegRead[24];
_IsoMon_DeviceSignals.voltageL2L3.bytes[3] := _RegRead[21];
_IsoMon_DeviceSignals.voltageL2L3.bytes[4] := _RegRead[22];

// 0x200C: voltageL1PE
_IsoMon_DeviceSignals.voltageL1PE.bytes[1] := _RegRead[27];
_IsoMon_DeviceSignals.voltageL1PE.bytes[2] := _RegRead[28];
_IsoMon_DeviceSignals.voltageL1PE.bytes[3] := _RegRead[25];
_IsoMon_DeviceSignals.voltageL1PE.bytes[4] := _RegRead[26];

// 0x200E: voltageL2PE
_IsoMon_DeviceSignals.voltageL2PE.bytes[1] := _RegRead[31];
_IsoMon_DeviceSignals.voltageL2PE.bytes[2] := _RegRead[32];
_IsoMon_DeviceSignals.voltageL2PE.bytes[3] := _RegRead[29];
_IsoMon_DeviceSignals.voltageL2PE.bytes[4] := _RegRead[30];

// 0x2010: voltageL3PE
_IsoMon_DeviceSignals.voltageL3PE.bytes[1] := _RegRead[35];
_IsoMon_DeviceSignals.voltageL3PE.bytes[2] := _RegRead[36];
_IsoMon_DeviceSignals.voltageL3PE.bytes[3] := _RegRead[33];
_IsoMon_DeviceSignals.voltageL3PE.bytes[4] := _RegRead[34];

// 0x2012: systemFrequency
_IsoMon_DeviceSignals.systemFrequency.bytes[1] := _RegRead[39];
_IsoMon_DeviceSignals.systemFrequency.bytes[2] := _RegRead[40];
_IsoMon_DeviceSignals.systemFrequency.bytes[3] := _RegRead[37];
_IsoMon_DeviceSignals.systemFrequency.bytes[4] := _RegRead[38];

// 0x2014: couplingToSystem
_IsoMon_DeviceSignals.couplingToSystem.bytes[1] := _RegRead[43];
_IsoMon_DeviceSignals.couplingToSystem.bytes[2] := _RegRead[44];
_IsoMon_DeviceSignals.couplingToSystem.bytes[3] := _RegRead[41];
_IsoMon_DeviceSignals.couplingToSystem.bytes[4] := _RegRead[42];

// 0x2016: couplingToEarth
_IsoMon_DeviceSignals.couplingToEarth.bytes[1] := _RegRead[47];
_IsoMon_DeviceSignals.couplingToEarth.bytes[2] := _RegRead[48];
_IsoMon_DeviceSignals.couplingToEarth.bytes[3] := _RegRead[45];
_IsoMon_DeviceSignals.couplingToEarth.bytes[4] := _RegRead[46];

// 0x2018: deviceError
_IsoMon_DeviceSignals.deviceError.bytes[1] := _RegRead[51];
_IsoMon_DeviceSignals.deviceError.bytes[2] := _RegRead[52];
_IsoMon_DeviceSignals.deviceError.bytes[3] := _RegRead[49];
_IsoMon_DeviceSignals.deviceError.bytes[4] := _RegRead[50];

// 0x201A: deviceInactive
_IsoMon_DeviceSignals.deviceInactive.bytes[1] := _RegRead[55];
_IsoMon_DeviceSignals.deviceInactive.bytes[2] := _RegRead[56];
_IsoMon_DeviceSignals.deviceInactive.bytes[3] := _RegRead[53];
_IsoMon_DeviceSignals.deviceInactive.bytes[4] := _RegRead[54];

// 0x201C: dcOffset
_IsoMon_DeviceSignals.dcOffset.bytes[1] := _RegRead[59];
_IsoMon_DeviceSignals.dcOffset.bytes[2] := _RegRead[60];
_IsoMon_DeviceSignals.dcOffset.bytes[3] := _RegRead[57];
_IsoMon_DeviceSignals.dcOffset.bytes[4] := _RegRead[58];

// 0x201E: measurementQuality
_IsoMon_DeviceSignals.measurementQuality.bytes[1] := _RegRead[63];
_IsoMon_DeviceSignals.measurementQuality.bytes[2] := _RegRead[64];
_IsoMon_DeviceSignals.measurementQuality.bytes[3] := _RegRead[61];
_IsoMon_DeviceSignals.measurementQuality.bytes[4] := _RegRead[62];

// 0x2020: symmetricalAlarm
_IsoMon_DeviceSignals.symmetricalAlarm.bytes[1] := _RegRead[67];
_IsoMon_DeviceSignals.symmetricalAlarm.bytes[2] := _RegRead[68];
_IsoMon_DeviceSignals.symmetricalAlarm.bytes[3] := _RegRead[65];
_IsoMon_DeviceSignals.symmetricalAlarm.bytes[4] := _RegRead[66];

// 0x2022: dcMinusAlarm
_IsoMon_DeviceSignals.dcMinusAlarm.bytes[1] := _RegRead[71];
_IsoMon_DeviceSignals.dcMinusAlarm.bytes[2] := _RegRead[72];
_IsoMon_DeviceSignals.dcMinusAlarm.bytes[3] := _RegRead[69];
_IsoMon_DeviceSignals.dcMinusAlarm.bytes[4] := _RegRead[70];

// 0x2024: dcPlusAlarm
_IsoMon_DeviceSignals.dcPlusAlarm.bytes[1] := _RegRead[75];
_IsoMon_DeviceSignals.dcPlusAlarm.bytes[2] := _RegRead[76];
_IsoMon_DeviceSignals.dcPlusAlarm.bytes[3] := _RegRead[73];
_IsoMon_DeviceSignals.dcPlusAlarm.bytes[4] := _RegRead[74];

// 0x2026: durationMeasuringPulse
_IsoMon_DeviceSignals.durationMeasuringPulse.bytes[1] := _RegRead[79];
_IsoMon_DeviceSignals.durationMeasuringPulse.bytes[2] := _RegRead[80];
_IsoMon_DeviceSignals.durationMeasuringPulse.bytes[3] := _RegRead[77];
_IsoMon_DeviceSignals.durationMeasuringPulse.bytes[4] := _RegRead[78];

// 0x2028: voltageDCPE
_IsoMon_DeviceSignals.voltageDCPE.bytes[1] := _RegRead[83];
_IsoMon_DeviceSignals.voltageDCPE.bytes[2] := _RegRead[84];
_IsoMon_DeviceSignals.voltageDCPE.bytes[3] := _RegRead[81];
_IsoMon_DeviceSignals.voltageDCPE.bytes[4] := _RegRead[82];
END_METHOD

METHOD PRIVATE cmdReadRegisters : BOOL
VAR_INPUT
END_VAR

VAR

END_VAR
CASE _RegReadState OF 
	0:
		IF (_modbus_IF.ReadRegisters.bBusy = FALSE) THEN
			_modbus_IF.ReadRegisters.nQuantity := SIZEOF(_RegRead)/2;
			_modbus_IF.ReadRegisters.cbLength  := SIZEOF(_RegRead);
			_modbus_IF.ReadRegisters.pDestAddr := ADR(_RegRead);
			_modbus_IF.ReadRegisters.nMBAddr   := 8192;
			_modbus_IF.ReadRegisters.bExecute  := TRUE;
			_RegReadState := 1;
		END_IF
	1:
		IF _modbus_IF.ReadRegisters.bBusy = TRUE THEN
			_modbus_IF.ReadRegisters.bExecute := FALSE;
			_RegReadState := 2;
		END_IF
	2:
		IF _modbus_IF.ReadRegisters.bBusy = FALSE THEN
			// A failed read used to go unnoticed: the HMI kept showing the last insulation
			// resistance with no fault. Now it faults (latched until reset) and the old values
			// are not re-parsed; stsCommOK says whether the readings are current.
			IF _modbus_IF.ReadRegisters.bError THEN
				_commOK := FALSE;
				setFault(1, 'Comms. Read Fault - insulation readings are not current');
			ELSE
				_commOK := TRUE;
				cmdParseRegisters();
			END_IF
			_RegReadState := 900;
		END_IF
END_CASE
END_METHOD

METHOD cmdReset : BOOL
setFault(0,'');
END_METHOD

METHOD PUBLIC cmdResetTrip : BOOL
VAR_INPUT

END_VAR
_cmdResetTrip := TRUE;
END_METHOD

METHOD PUBLIC cmdTest : BOOL
VAR_INPUT
	IO_value	: BOOL;
END_VAR
IF IO_OUT_Test <> 0 THEN
	IO_OUT_Test^ := IO_value;
END_IF
END_METHOD

METHOD PRIVATE FaultHandler : BOOL
VAR_INPUT
END_VAR
IF IO_IN_DeviceTrip^ = FALSE THEN
	setFault(1,'Loss of isolation between HVDC and ground');
END_IF

IF IO_IN_DeviceWarning^ = FALSE THEN
	sendWarning('Isolation Warning - abnormally low isolation to ground',1);
END_IF
END_METHOD

(*FB_Init is always available implicitly and it is used primarily for initialization.
The return value is not evaluated. For a specific influence, you can also declare the
methods explicitly and provide additional code there with the standard initialization
code. You can evaluate the return value.*)
METHOD FB_Init : BOOL
VAR_INPUT
	(* TRUE: the retain variables are initialized (reset warm / reset cold)*)
	bInitRetains	: BOOL;
	(* TRUE: the instance will be copied to the copy code afterward (online change)   *)
	bInCopyCode	: BOOL;
	cfgDeviceName	: STRING;
	cfgEnable	: BOOL;
	cfgInitEventClass	: BOOL;
END_VAR
THIS^.cfgDeviceName 		:= 		cfgDeviceName; 		
THIS^.cfgEnable 			:= 	    cfgEnable; 	
THIS^.cfgInitEventClass		:= 		cfgInitEventClass;
END_METHOD

METHOD updateHMI : BOOL
VAR_INPUT
END_VAR
HMI_deviceSignals.insulationResistance_kOhm := _isoMon_DeviceSignals.insulationResistance.value / 1000;
HMI_deviceSignals.minInsulationValue		:= _isoMon_DeviceSignals.minInsulationValue.value / 1000;
HMI_deviceSignals.voltageDCPlusToMinus		:= _isoMon_DeviceSignals.voltageL1L3.value;
HMI_deviceSignals.voltageDCPlusToPE			:= _isoMon_DeviceSignals.voltageL1PE.value;
HMI_deviceSignals.voltageDCMinusToPE		:= _isoMon_DeviceSignals.voltageL3PE.value;
HMI_deviceSignals.couplingToSystem			:= _isoMon_DeviceSignals.couplingToSystem.value;
HMI_deviceSignals.couplingtoEarth			:= _isoMon_DeviceSignals.couplingToEarth.value;
HMI_deviceSignals.deviceError				:= _isoMon_DeviceSignals.deviceError.value;
HMI_deviceSignals.deviceInactive			:= _isoMon_DeviceSignals.deviceInactive.value;
HMI_deviceSignals.dcOffset					:= _isoMon_DeviceSignals.dcOffset.value;
HMI_deviceSignals.measurementQuality		:= _isoMon_DeviceSignals.measurementQuality.value;
HMI.HMIbaseDevice := HMIbaseDevice;

//Reset command from HMI
IF HMI.ocmdTripReset OR inpReset OR _cmdResetTrip THEN
	TOFResetTrig 		:= TRUE;
	HMI.ocmdTripReset	:= FALSE;
	_cmdResetTrip		:= FALSE;
END_IF

IF TOFReset.Q THEN
	IO_OUT_TripReset^ := TRUE;
	TOFResetTrig	  := FALSE;
ELSE
	IO_OUT_TripReset^ := FALSE;
END_IF

//Test command from HMI
IF HMI.ocmdTest THEN
	TOFTestTrig			:= TRUE;
	HMI.ocmdTest		:= FALSE;
END_IF

IF TOFTest.Q THEN
	IO_OUT_Test^	  := TRUE;
	TOFTestTrig		  := FALSE;
ELSE
	IO_OUT_Test^	  := FALSE;
END_IF
END_METHOD

END_FUNCTION_BLOCK

// ---- POUs/FBs/Devices/fb_Dev_Machine.TcPOU
FUNCTION_BLOCK fb_Dev_Machine EXTENDS abs_fb_Device

VAR_INPUT
	start				: BOOL;
	stop				: BOOL;
	SafetyPowerOn		: BOOL;
	SafetyFaultActive	: BOOL;
END_VAR

DeviceLogic();
Interlock.name := _DeviceName;
Interlock(inpConfig := _dataInterlock);


faultHandler();

METHOD cmdReset : BOOL
IF stsFaulted THEN
	setFault(0,'');
END_IF
END_METHOD

METHOD faultHandler : BOOL
VAR_INPUT
END_VAR
IF stop THEN
	sendWarning('Machine STOP pressed',1);
END_IF

IF inpReset THEN
	sendLog('Machine RESET', 1);
ELSE
	_logChannels[1] := '';
END_IF

IF start THEN
	sendLog('Auto sequence started', 2);
ELSE
	_logChannels[2] := '';
END_IF

IF _inAuto THEN
	sendLog('Machine set to AUTO',3);
ELSE
	sendLog('Machine set to MANUAL',3);
END_IF

IF safetyPowerOn THEN
	sendLog('Safety - Power ON', 4);
ELSE
	sendLog('Safety - Power OFF', 4);
END_IF
END_METHOD

END_FUNCTION_BLOCK

// ---- POUs/FBs/Devices/fb_Dev_PSU_ITECH.TcPOU
(*
    fb_Dev_PSU_ITECH — ITECH programmable DC supply (IT6000 / IT6600C) over Modbus TCP.

    All traffic goes through fb_Modbus_Driver: one connection, requests strictly in series,
    a pause of the type's scan time between transactions (these supplies are slow and do not
    like to be rushed).

    COMMS LATCH. The FIRST failed read or write stops ALL traffic to the supply — no retries,
    no reconnect loop — and raises a fault. Nothing is sent again until a reset (inpReset,
    an HMI reset, or cmdReset()). ITECHs misbehave when they are polled while they are
    refusing requests, so the block waits for a person rather than hammering them.

    BASELINE BEFORE WRITE. After every (re)start the block reads the supply's current settings
    first and seeds its command image from them; writes are held until then, so a restart
    never sends zeros or stale setpoints. When the restart follows a comms fault, the output
    is commanded OFF as part of that baseline: the PLC lost sight of the supply, so an
    operator re-enables it deliberately. A reset never re-energises anything.

    Usage:
        PSU1 : fb_Dev_PSU_ITECH(cfgDeviceName := 'PSU1', cfgEnable := TRUE, cfgInitEventClass := TRUE);
        PSU1.cfgModbusConfig := cfg;        // IP, port (0 = 502), unit id, timeout (0 = 1 s)
        PSU1(ITECH_Type := 'IT6600C', IOIn_OKToUnInhibit := ..., IOOut_Inhibit := ADR(...));
*)
FUNCTION_BLOCK fb_Dev_PSU_ITECH EXTENDS abs_fb_Device
VAR_INPUT
    ITECH_Type          : STRING;           // 'IT6600C' or 'IT6000'
    IOIn_OKToUnInhibit  : BOOL;
    IOOut_Inhibit       : POINTER TO BOOL;
END_VAR

VAR_OUTPUT
    stsDCSourceState    : UDINT;
    stsDCMode           : UDINT;
    stsDCSource_V_SP    : REAL;
    stsDCMeterV         : REAL;
    stsDCMeterI         : REAL;
    stsDCMeterP         : REAL;
    stsCommFaulted      : BOOL;             // comms stopped by the latch; cleared by a reset
END_VAR

VAR PERSISTENT
    HMI_DeviceSignals   : ST_ITECH_HMI_DeviceSignals;
END_VAR

VAR
    // Modbus — all comms go through the driver
    _modbus_cfg         : ST_Modbus_Device_Config;
    _mb                 : fb_Modbus_Driver;
    _arrReadConfig      : ARRAY[1..47] OF ST_MBSignalConfig;
    _arrReadResults     : ARRAY[1..47] OF ST_MBReadResult;
    _arrWriteConfig     : ARRAY[1..34] OF ST_MBSignalConfig;
    _arrWriteData       : ARRAY[1..34] OF ST_MBWriteData;
    // one-shot protection-reset write (a register that must NOT be written every cycle)
    _mbReset            : fb_Modbus_Driver;
    _arrResetConfig     : ARRAY[1..1] OF ST_MBSignalConfig;
    _arrResetData       : ARRAY[1..1] OF ST_MBWriteData;

    // register map of the selected type
    _mapValid           : BOOL;
    _hasExtStatus       : BOOL;             // IT6600C publishes 8 system-status values, IT6000 two
    _scanTime           : TIME;
    _regDCMeter         : UINT;
    _regDCSource        : UINT;
    _regSystemStatus    : UINT;
    _regProtection      : UINT;
    _regSoftwareFaults  : UINT;
    _regOnOff           : UINT;
    _regResetFault      : UINT;
    _activeType         : STRING;
    _mapChanged         : BOOL;

    // comms state
    _commRun            : BOOL;
    _commRunPrev        : BOOL;
    _commFaulted        : BOOL;
    _commFaultSeen      : BOOL;             // set by the latch; the next baseline commands OFF
    _baselineTaken      : BOOL;
    _readCount          : UINT;
    _lastReadCycles     : UDINT;
    _wdTime             : TIME;
    _tonReadWatchdog    : TON;
    _resetCalled        : BOOL;
    _resetTrig          : R_TRIG;
    _deviceResetPending : BOOL;
    _resetRun           : BOOL;
    _resetRunPrev       : BOOL;
    _baselineCurrentLimit : REAL := 20.5;

    // device images
    _device             : ST_ITECH_DeviceSignals;   // what the supply reports
    _command            : ST_ITECH_DeviceSignals;   // what this block writes
    _swFaultReg         : UDINT;
    _SoftwareFaults     : ST_ITECH_SoftwareFaults;
    _DeviceFaults       : ST_ITECH_QuestionRegister;
END_VAR

VAR CONSTANT
    // read table layout (index offsets into _arrReadConfig / _arrReadResults)
    cRD_METER           : UINT := 0;    // 1..6    DC meter
    cRD_SOURCE          : UINT := 6;    // 7..21   DC source
    cRD_PROT            : UINT := 21;   // 22..38  protection
    cRD_SWF             : UINT := 39;   // 39      software faults
    cRD_SYS             : UINT := 39;   // 40..47  system status (IT6000: 40..41 only)
    // write table layout
    cWR_ONOFF           : UINT := 0;    // 1..2    on/off (two 16-bit registers, see writeImage)
    cWR_SOURCE          : UINT := 2;    // 3..17   DC source
    cWR_PROT            : UINT := 17;   // 18..34  protection
END_VAR

DeviceLogic();
setInterlock();

IF IOOut_Inhibit <> 0 THEN
    IOOut_Inhibit^ := IOIn_OKToUnInhibit;
END_IF

selectRegisterMap();

IF _enabled THEN
    FaultHandler();
    IF _baselineTaken THEN
        setCommandValues();
    END_IF
END_IF

runComms();

IF _baselineTaken AND NOT _commFaulted THEN
    setStatusValues();
END_IF

stsCommFaulted := _commFaulted;
updateHMI();

// Current limit applied as +/- to the command image when it is seeded from the supply
// after a (re)start. Default 20.5 A (the value this block has always applied); 0 = keep the
// supply's own limits.
PROPERTY cfgBaselineCurrentLimit : REAL
GET
cfgBaselineCurrentLimit := _baselineCurrentLimit;
END_GET
SET
_baselineCurrentLimit := cfgBaselineCurrentLimit;
END_SET
END_PROPERTY

PROPERTY cfgModbusConfig : ST_Modbus_Device_Config
GET
cfgModbusConfig := _modbus_cfg;
END_GET
SET
// Applied the next time comms (re)start (enable, reset after a comms fault, type change).
_modbus_cfg := cfgModbusConfig;
END_SET
END_PROPERTY

METHOD PRIVATE checkDeviceFaults : BOOL
IF _DeviceFaults.overVoltageProtection THEN
    setFault(1, 'Internal Fault - Overvoltage protection');
END_IF
IF _DeviceFaults.overCurrentProtection THEN
    setFault(1, 'Internal Fault - Overcurrent protection');
END_IF
IF _DeviceFaults.overPowerProtection THEN
    setFault(1, 'Internal Fault - Overpower protection');
END_IF
IF _DeviceFaults.underVoltageProtection THEN
    setFault(1, 'Internal Fault - Undervoltage protection');
END_IF
IF _DeviceFaults.overTempProtection THEN
    setFault(1, 'Internal Fault - Overtemperature protection');
END_IF
IF _DeviceFaults.underCurrentProtection THEN
    setFault(1, 'Internal Fault - Undercurrent protection');
END_IF
IF _DeviceFaults.senseFault THEN
    setFault(1, 'Internal Fault - Sense fault');
END_IF
IF _DeviceFaults.currentSharingFault THEN
    setFault(1, 'Internal Fault - Current sharing fault');
END_IF
IF _DeviceFaults.externalInhibit THEN
    setFault(1, 'Device inhibited');
END_IF
IF _DeviceFaults.faultProtection THEN
    setFault(1, 'Internal Fault - Device fault protection active');
END_IF
IF _DeviceFaults.loopOscFailure THEN
    setFault(1, 'Internal Fault - Loop oscillation failure');
END_IF
IF _DeviceFaults.outputNotRegulated THEN
    setFault(1, 'Internal Fault - Output not regulated');
END_IF

IF _SoftwareFaults.outputReverseProtection THEN
    sendWarning('Output reverse protection', 10);
END_IF
IF _SoftwareFaults.multiMasterUnitsAbnormal THEN
    sendWarning('Multimaster unit abnormal', 11);
END_IF
IF _SoftwareFaults.opticalFiberUnlocked_singleMaster THEN
    sendWarning('Optical fiber NOK', 12);
END_IF
IF _SoftwareFaults.moduleCheckingFailure THEN
    sendWarning('Inconsistent master and slave module parameters', 13);
END_IF
IF _SoftwareFaults.unevenCurrentProtection THEN
    sendWarning('Uneven current protection', 14);
END_IF
IF _SoftwareFaults.masterUnitPowerFailureProtection THEN
    sendWarning('Master unit power failure protection', 15);
END_IF
IF _SoftwareFaults.capacitorOverCurrentprotection THEN
    sendWarning('Capacitor overcurrent protection', 16);
END_IF
IF _SoftwareFaults.slaveUnitPowerFailureProtection THEN
    sendWarning('Slave unit power failure protection', 17);
END_IF
END_METHOD

METHOD cmdDCSourceEnable : BOOL
VAR_INPUT
    onRequest   : BOOL;
END_VAR
IF onRequest THEN
    _command.System.ON_OFF := 1;
ELSE
    _command.System.ON_OFF := 0;
    HMI_DeviceSignals.deviceSignals_write.System.ON_OFF := 0;
END_IF
END_METHOD

METHOD cmdReset : BOOL
// Called every scan while inpReset is held (abs_fb_Device.DeviceLogic); runComms acts on the
// rising edge only, so holding reset does not turn into a retry loop against the supply.
IF stsFaulted THEN
    setFault(0, '');
END_IF
_resetCalled := TRUE;
END_METHOD

METHOD cmdSetCurrentLimits : BOOL
VAR_INPUT
    currentLimitHigh : REAL;
    currentLimitLow  : REAL;
END_VAR
_command.DCSource.DCCurrentHigh := currentLimitHigh;
_command.DCSource.DCCurrentLow  := currentLimitLow;
END_METHOD

METHOD PUBLIC cmdSetVoltageSP : BOOL
VAR_INPUT
    voltageSP   : REAL;
END_VAR
_command.DCSource.DCVoltSP := voltageSP;
END_METHOD

METHOD PRIVATE configureDriver : BOOL
VAR
    _timeout    : TIME;
    _port       : UINT;
    _i          : UINT;
END_VAR
// Called on the scan comms (re)start, BEFORE the enable edge reaches the driver: the driver
// only accepts properties while it is not initialised.
_timeout := _modbus_cfg.cfgTimeout;
IF _timeout = T#0S THEN
    _timeout := T#1S;
END_IF
_port := _modbus_cfg.cfgTCPPort;
IF _port = 0 THEN
    _port := 502;
END_IF

_mb.ipAddress            := _modbus_cfg.cfgIP_address;
_mb.port                 := _port;
_mb.unitId               := _modbus_cfg.cfgUnitID;
_mb.timeout              := _timeout;
_mb.pollInterval         := _scanTime;
_mb.commandDelay         := _scanTime;      // pause between transactions, as these supplies need
_mb.writeCycleInterval   := _scanTime;
_mb.wordOrder            := E_WordOrder.BigEndian;
// This block latches on the FIRST failure itself; keep the driver's own retry logic out of the way.
_mb.maxConsecFails       := 1000;
_mb.maxReconnectAttempts := 1000;
_mb.staleThreshold       := T#10S;

// ── reads ──────────────────────────────────────────────────────────────────────────────────
// DC meter
setRead(cRD_METER + 1,  _regDCMeter + 0,  TRUE);    // Vrms
setRead(cRD_METER + 2,  _regDCMeter + 2,  TRUE);    // Irms
setRead(cRD_METER + 3,  _regDCMeter + 4,  TRUE);    // Prms (IT6000: kW, IT6600C: W)
setRead(cRD_METER + 4,  _regDCMeter + 6,  FALSE);   // operation register
setRead(cRD_METER + 5,  _regDCMeter + 8,  FALSE);   // state register
setRead(cRD_METER + 6,  _regDCMeter + 10, FALSE);   // questionable register
// DC source
setRead(cRD_SOURCE + 1,  _regDCSource + 0,  FALSE); // mode
setRead(cRD_SOURCE + 2,  _regDCSource + 2,  TRUE);  // voltage SP
setRead(cRD_SOURCE + 3,  _regDCSource + 4,  TRUE);  // voltage rise
setRead(cRD_SOURCE + 4,  _regDCSource + 6,  TRUE);  // voltage fall
setRead(cRD_SOURCE + 5,  _regDCSource + 8,  TRUE);  // current SP
setRead(cRD_SOURCE + 6,  _regDCSource + 10, TRUE);  // current rise
setRead(cRD_SOURCE + 7,  _regDCSource + 12, TRUE);  // current fall
setRead(cRD_SOURCE + 8,  _regDCSource + 14, TRUE);  // voltage high
setRead(cRD_SOURCE + 9,  _regDCSource + 16, TRUE);  // voltage low
setRead(cRD_SOURCE + 10, _regDCSource + 18, TRUE);  // current high
setRead(cRD_SOURCE + 11, _regDCSource + 20, TRUE);  // current low
setRead(cRD_SOURCE + 12, _regDCSource + 22, FALSE); // CC speed state
setRead(cRD_SOURCE + 13, _regDCSource + 24, FALSE); // CV speed state
setRead(cRD_SOURCE + 14, _regDCSource + 26, TRUE);  // power high
setRead(cRD_SOURCE + 15, _regDCSource + 28, TRUE);  // power low
// protection: OVP, OCP, OPP (state, level, delay), UCP, UVP (state, level, delay, warm-up)
FOR _i := 0 TO 2 DO
    setRead(cRD_PROT + 1 + _i * 3, _regProtection + _i * 6 + 0, FALSE);
    setRead(cRD_PROT + 2 + _i * 3, _regProtection + _i * 6 + 2, TRUE);
    setRead(cRD_PROT + 3 + _i * 3, _regProtection + _i * 6 + 4, TRUE);
END_FOR
FOR _i := 0 TO 1 DO
    setRead(cRD_PROT + 10 + _i * 4, _regProtection + 18 + _i * 8 + 0, FALSE);
    setRead(cRD_PROT + 11 + _i * 4, _regProtection + 18 + _i * 8 + 2, TRUE);
    setRead(cRD_PROT + 12 + _i * 4, _regProtection + 18 + _i * 8 + 4, TRUE);
    setRead(cRD_PROT + 13 + _i * 4, _regProtection + 18 + _i * 8 + 6, TRUE);
END_FOR
// software faults
setRead(cRD_SWF, _regSoftwareFaults, FALSE);
// system status
setRead(cRD_SYS + 1, _regSystemStatus + 0, FALSE);  // on/off
setRead(cRD_SYS + 2, _regSystemStatus + 2, TRUE);   // sense voltage
IF _hasExtStatus THEN
    setRead(cRD_SYS + 3, _regSystemStatus + 4,  FALSE); // heartbeat
    setRead(cRD_SYS + 4, _regSystemStatus + 6,  FALSE); // timer on/off
    setRead(cRD_SYS + 5, _regSystemStatus + 8,  FALSE); // remote sense status
    setRead(cRD_SYS + 6, _regSystemStatus + 10, TRUE);  // remote sense level
    setRead(cRD_SYS + 7, _regSystemStatus + 12, FALSE); // output R zero
    setRead(cRD_SYS + 8, _regSystemStatus + 14, FALSE); // measure cycle
    _readCount := cRD_SYS + 8;
ELSE
    _readCount := cRD_SYS + 2;
END_IF
_mb.readSignalCount := _readCount;

// ── writes ─────────────────────────────────────────────────────────────────────────────────
_arrWriteConfig[cWR_ONOFF + 1].modbusAddr := 400001 + UINT_TO_UDINT(_regOnOff);
_arrWriteConfig[cWR_ONOFF + 1].dataType   := E_MBDataType.mbUInt16;
_arrWriteConfig[cWR_ONOFF + 2].modbusAddr := 400001 + UINT_TO_UDINT(_regOnOff) + 1;
_arrWriteConfig[cWR_ONOFF + 2].dataType   := E_MBDataType.mbUInt16;
FOR _i := 1 TO 15 DO
    // same 15 values, same order and types as the DC-source read block
    setWrite(cWR_SOURCE + _i, _regDCSource + (_i - 1) * 2,
             _arrReadConfig[cRD_SOURCE + _i].dataType = E_MBDataType.mbReal32);
END_FOR
FOR _i := 1 TO 17 DO
    setWrite(cWR_PROT + _i, _regProtection + (_i - 1) * 2,
             _arrReadConfig[cRD_PROT + _i].dataType = E_MBDataType.mbReal32);
END_FOR
_mb.writeSignalCount := cWR_PROT + 17;

FOR _i := 1 TO cWR_PROT + 17 DO
    _arrWriteData[_i].writeError   := FALSE;
    _arrWriteData[_i].writeSuccess := FALSE;
END_FOR

// watchdog on read-cycle progress: generous against a normal cycle, short against a stuck one
_wdTime := MAX(T#5S, UDINT_TO_TIME(6 * TIME_TO_UDINT(_scanTime + _timeout)));
_activeType := ITECH_Type;
END_METHOD

METHOD PRIVATE deviceResetWrite : BOOL
// The supply clears its latched protection on a write to the reset register (value 0, as it
// always was). It must be written ONCE per reset, never on every write cycle, so it gets its
// own driver instance that runs only while a reset is pending.
_resetRun := _deviceResetPending AND _baselineTaken AND NOT _commFaulted;

IF _resetRun AND NOT _resetRunPrev THEN
    _mbReset.ipAddress            := _mb.ipAddress;
    _mbReset.port                 := _mb.port;
    _mbReset.unitId               := _mb.unitId;
    _mbReset.timeout              := _mb.timeout;
    _mbReset.pollInterval         := T#1S;
    _mbReset.commandDelay         := _scanTime;
    _mbReset.writeCycleInterval   := T#10MS;
    _mbReset.wordOrder            := E_WordOrder.BigEndian;
    _mbReset.maxConsecFails       := 1000;
    _mbReset.maxReconnectAttempts := 1000;
    _mbReset.readSignalCount      := 0;
    _mbReset.writeSignalCount     := 1;
    _arrResetConfig[1].modbusAddr := 400001 + UINT_TO_UDINT(_regResetFault);
    _arrResetConfig[1].dataType   := E_MBDataType.mbUInt32;
    _arrResetData[1].valueUdint   := 0;
    _arrResetData[1].writeError   := FALSE;
    _arrResetData[1].writeSuccess := FALSE;
END_IF
_resetRunPrev := _resetRun;

_mbReset(
    inpEnable           := _resetRun,
    inpPtrReadConfig    := 0,
    inpPtrReadResults   := 0,
    inpPtrWriteConfig   := ADR(_arrResetConfig),
    inpPtrWriteData     := ADR(_arrResetData));
_mbReset.cycle();

IF _resetRun THEN
    IF _arrResetData[1].writeError THEN
        latchCommFault('Modbus write failed (protection reset) - comms stopped until reset');
    ELSIF _arrResetData[1].writeSuccess THEN
        _deviceResetPending := FALSE;   // next scan disables the one-shot driver
    END_IF
END_IF
END_METHOD

METHOD PRIVATE FaultHandler : BOOL
// Turn off if already on and the interlock drops
IF NOT(Interlock.outInterlockOK) AND stsDCSourceState = 1 THEN
    cmdDCSourceEnable(0);
    setFault(1, Interlock.stsFirstOut);
END_IF

// Short-circuit detection
IF stsDCSourceState = 1 AND stsDCMode = 1 THEN
    IF (stsDCMeterV - stsDCSource_V_SP) < 20 AND stsDCMeterI > 5 THEN
        setFault(1, 'Shortcircuit current detected');
    END_IF
END_IF

IF stsFaulted OR NOT(Interlock.outInterlockOK) THEN
    cmdDCSourceEnable(0);
    HMI_DeviceSignals.deviceSignals_write.System.ON_OFF := 0;
END_IF

IF NOT _mapValid THEN
    setFault(1, CONCAT('Unknown ITECH_Type: ', ITECH_Type));
END_IF

IF _baselineTaken AND NOT _commFaulted THEN
    parseFaults();
    checkDeviceFaults();
END_IF
END_METHOD

//FB_Init is always available implicitly and it is used primarily for initialization.
//The return value is not evaluated. For a specific influence, you can also declare the
//methods explicitly and provide additional code there with the standard initialization
//code. You can evaluate the return value.
METHOD FB_Init : BOOL
VAR_INPUT
    bInitRetains        : BOOL; // TRUE: the retain variables are initialized (reset warm / reset cold)
    bInCopyCode         : BOOL; // TRUE: the instance will be copied to the copy code afterward (online change)
    cfgDeviceName       : STRING;
    cfgEnable           : BOOL;
    cfgInitEventClass   : BOOL;
END_VAR
THIS^.cfgDeviceName     := cfgDeviceName;
THIS^.cfgEnable         := cfgEnable;
THIS^.cfgInitEventClass := cfgInitEventClass;
END_METHOD

METHOD PRIVATE initParameters : BOOL
// The operator's editable values start from what the supply is actually set to.
HMI_DeviceSignals.deviceSignals_write := _device;
END_METHOD

METHOD PRIVATE latchCommFault : BOOL
VAR_INPUT
    inpMessage  : STRING;
END_VAR
// Stop ALL traffic to the supply in THIS scan, before the driver can send anything else,
// and stay stopped until a reset.
_commFaulted := TRUE;
_commFaultSeen := TRUE;
setFault(1, inpMessage);

_mb(inpEnable := FALSE);
_mb.cycle();
_mbReset(inpEnable := FALSE);
_mbReset.cycle();

_commRunPrev        := FALSE;
_resetRunPrev       := FALSE;
_baselineTaken      := FALSE;
_deviceResetPending := FALSE;
_tonReadWatchdog(IN := FALSE);
END_METHOD

